(* IEC 61131-3 sources: NachHouse_TST/OSCAT_BasicLib/OscatBasicLib_333a (part 6) *)

(* ---- Device_Driver.ST ---- *)
(* @PATH := '\/Engineering\/automation' *)
FUNCTION_BLOCK DRIVER_1
(*
  driver_1 is a multi purpose driver.
  a rising edge on in sets the output high if toggle is flase. while toggle is true, a rising edge on in toggles the output Q.
  if a timeout is specified the output q will be reset to false automatically after the timeout has elapsed.
  a asynchronous reset and set will force the output high or low respectively.

  version 1.0 2 jan 2008
  programmer  hugo
  tested by   tobias
*)
  VAR_INPUT //???CONSTANT
    Toggle_Mode : BOOL;
    Timeout : TIME;
  END_VAR
  VAR_INPUT
    SET : BOOL;
    IN : BOOL;
    RST : BOOL;
  END_VAR
  VAR_OUTPUT
    Q : BOOL;
  END_VAR
  VAR
    off : TON;
    edge: BOOL;
  END_VAR

  IF off.Q THEN Q := FALSE; END_IF;
  IF rst THEN
    Q := FALSE;
  ELSIF set THEN
    Q := TRUE;
  ELSIF IN AND NOT edge THEN
    IF toggle_mode THEN q := NOT Q; ELSE q := TRUE; END_IF;
  END_IF;
  edge := in;
  IF timeout > t#0s THEN off(in := Q, PT := Timeout); END_IF;

(* revision history
  hm  2. jan 2008   rev 1.0
    original version
*)
END_FUNCTION_BLOCK

(* @PATH := '\/Engineering\/automation' *)
FUNCTION_BLOCK DRIVER_4
(*
  driver_4 is a 4 channel multi purpose driver.
  a rising edge on in? sets the output Q? high if toggle_mode is flase. while toggle_mode is true, a rising edge on in? toggles the output Q?.
  if a timeout is specified the output Q? will be reset to false automatically after the timeout has elapsed.
  a asynchronous reset and set will force the output high or low respectively.
  an asynchronous set will force all outputs high simultaneously

  version 1.0 2 jan 2008
  programmer  hugo
  tested by   tobias
*)
  VAR_INPUT //???CONSTANT
    Toggle_Mode : BOOL;
    Timeout : TIME;
  END_VAR
  VAR_INPUT
    SET : BOOL;
    IN0, IN1, IN2, IN3 : BOOL;
    RST : BOOL;
  END_VAR
  VAR_OUTPUT
    Q0, Q1, Q2, Q3 : BOOL;
  END_VAR
  VAR
    d0, d1, d2, d3 : DRIVER_1;
  END_VAR

  D0(Set:=set, in:=in0, rst:=rst, toggle_mode:=toggle_mode, timeout:=timeout);
  D1(Set:=set, in:=in1, rst:=rst, toggle_mode:=toggle_mode, timeout:=timeout);
  D2(Set:=set, in:=in2, rst:=rst, toggle_mode:=toggle_mode, timeout:=timeout);
  D3(Set:=set, in:=in3, rst:=rst, toggle_mode:=toggle_mode, timeout:=timeout);
  Q0 := D0.Q;
  Q1 := D1.Q;
  Q2 := D2.Q;
  Q3 := D3.Q;

(* revision history
  hm  2. jan 2008   rev 1.0
    original version
*)
END_FUNCTION_BLOCK

(* @PATH := '\/Engineering\/automation' *)
FUNCTION_BLOCK DRIVER_4C
(*
  driver_4C is a multi purpose driver.
  a rising edge on in switches from S0 state S1 and the next edge to state S2 and so on.
  in state S0 all outputs Q are FALSE.
  The stet of the Outputs in any state S? is configurable with setup variables.
  The variables S1..S5 define the states, while the sequence is terminated when a state Variable S? = 0.
  The lower bits 0..3 of the state vars S? are corresponding to the Outputs Q0..Q3

  version 1.0 23. mar. 2009
  programmer  hugo
  tested by tobias
*)
  VAR_INPUT
    IN : BOOL;
    RST : BOOL;
  END_VAR
  VAR_INPUT //??? CONSTANT
    Timeout : TIME;
    SX : ARRAY[1..7] OF BYTE := [1,3,7,15];
  END_VAR
  VAR_OUTPUT
    SN : INT;
    Q0 : BOOL;
    Q1 : BOOL;
    Q2 : BOOL;
    Q3 : BOOL;
  END_VAR
  VAR
    off : TON;
    edge: BOOL;
  END_VAR

  IF RST OR off.Q THEN
    SN := 0;
  ELSIF IN AND NOT edge THEN
    SN := SN + 1;
    IF SN > 7 OR SX[SN] = 0 THEN SN := 0; END_IF;
  END_IF;
  edge := in;
  IF SN > 0 THEN
    Q0 := SX[SN].0;
    Q1 := SX[SN].1;
    Q2 := SX[SN].2;
    Q3 := SX[SN].3;
  ELSE
    Q0 := FALSE;
    Q1 := FALSE;
    Q2 := FALSE;
    Q3 := FALSE;
  END_IF;

  (* maximaum timeout *)
  IF timeout > t#0s THEN off(in := SN > 0, PT := Timeout); END_IF;

(* revision history
  hm  23. mar. 2009 rev 1.0
    original version
*)
END_FUNCTION_BLOCK

(* @PATH := '\/Engineering\/automation' *)
FUNCTION_BLOCK FLOW_CONTROL
(*
  FLOW_CONTROL switches a valves depending on the input in.
  flow control also limits the maximum ontime of the valve and controls pressure on the output side.

  version 1.0 28. jun. 2008
  programmer  hugo
  tested by oscat
*)
  VAR_INPUT
    IN : BOOL;
    REQ : BOOL;
    ENQ : BOOL;
    RST : BOOL;
  END_VAR
  VAR_INPUT //???CONSTANT
    T_AUTO : TIME := T#1h;
    T_DELAY : TIME := T#23h;
  END_VAR
  VAR_OUTPUT
    Q : BOOL;
    STATUS : BYTE;
  END_VAR
  VAR
    timer : TP_1D;
  END_VAR

  STATUS := 100;
  IF RST THEN
    Q := FALSE;
    timer(rst := TRUE);
    timer.RST := FALSE;
    STATUS := 103;
  ELSIF ENQ THEN
    IF IN THEN
      status := 101;
    END_IF;
    IF REQ THEN
      (* timer will generate a timed pulse after TP goes high *)
      timer.PT1 := T_AUTO;
      timer.PTD := T_DELAY;
      timer.IN := TRUE;
      STATUS := 102;
    END_IF;
  END_IF;

  (* set output and run timer *)
  timer();
  timer.IN := FALSE;
  Q := (IN AND ENQ) OR timer.Q;

(* revision history
  hm  28. jun. 2008   rev 1.0
    original version
*)
END_FUNCTION_BLOCK

(* @PATH := '\/Engineering\/automation' *)
FUNCTION_BLOCK FT_Profile
(*
  FT_Profile generates an output signal which is defined by values over a time scale.
  the different values are connected by ramps between the individual values.
  a rising edge on E starts the output signal generation and E = True can delay time_3 / value_3 as long as it stays true.
  an additional multiplier K can be used to multiply the output and an offset O can be added to the output dynamically.

  version 1.1 15 sep 2007
  programmer  tobias
  tested by   hugo
*)
  VAR_INPUT
    K : REAL := 1.0;
    O : REAL;
    M : REAL := 1.0;
    E : BOOL;
  END_VAR
  VAR_INPUT //???CONSTANT
    value_0 : REAL;
    time_1 : TIME;
    value_1 : REAL;
    time_2 : TIME;
    value_2 : REAL;
    time_3 : TIME;
    value_3 : REAL;
    time_10 : TIME;
    value_10 : REAL;
    time_11 : TIME;
    value_11 : REAL;
    time_12 : TIME;
    value_12 : REAL;
    time_13 : TIME;
    value_13 : REAL;
  END_VAR
  VAR_OUTPUT
    Y : REAL;
    RUN : BOOL;
    ET : TIME;
  END_VAR
  VAR
    tx : TIME;
    edge : BOOL;
    state: BYTE;
    ta: TIME;
    tb: TIME;
    t0 : TIME;
    temp: REAL;
    va: REAL;
    vb: REAL;
  END_VAR

  (* read system time *)
  tx := DWORD_TO_TIME(T_PLC_MS());

  (* determine start condition *)
  IF E AND NOT edge THEN
    RUN := TRUE;
    ET := t#0s;
    t0 := tx;
    ta := tx;
    tb := multime(time_1, M);
    va := value_0;
    vb := value_1;
    temp := value_0;
    state := 1;
  END_IF;
  edge := E;

  (* generate startup profile *)
  IF run THEN
    CASE BYTE_TO_USINT(state) OF
      1:  IF tx - ta >= tb THEN
          ta := ta + tb;
          tb := multime(time_2 - time_1, M);
          va := value_1;
          vb := value_2;
          temp := value_1;
          state := 2;
        ELSE
          temp := ((vb - va) * TIME_TO_REAL(tx - ta) / TIME_TO_REAL(tb) + va);
        END_IF;
      2:  IF tx - ta >= tb THEN
          ta := ta + tb;
          tb := multime(time_3 - time_2, M);
          va := value_2;
          vb := value_3;
          temp := value_2;
          state := 3;
        ELSE
          temp := ((vb - va) * TIME_TO_REAL(tx - ta) / TIME_TO_REAL(tb) + va);
        END_IF;
      3:  IF tx - ta >= tb THEN
          ta := ta + tb;
          tb := multime(time_10 - time_3, M);
          va := value_3;
          vb := value_10;
          temp := value_3;
          state := 4;
        ELSE
          temp := ((vb - va) * TIME_TO_REAL(tx - ta) / TIME_TO_REAL(tb) + va);
        END_IF;
      4 : IF tx - ta >= tb THEN
          ta := ta + tb;
          tb := multime(time_11 - time_10, M);
          va := value_10;
          vb := value_11;
          temp := value_10;
          IF E THEN state := 5; ELSE state := 6; END_IF;
        ELSE
          temp := ((vb - va) * TIME_TO_REAL(tx - ta) / TIME_TO_REAL(tb) + va);
        END_IF;
      5:  (* extend the signal while E is true *)
        IF E THEN
          ta := tx;
        ELSE
          state := 6;
        END_IF;
      6:  IF tx - ta >= tb THEN
          ta := ta + tb;
          tb := multime(time_12 - time_11, M);
          va := value_11;
          vb := value_12;
          temp := value_11;
          state := 7;
        ELSE
          temp := ((vb - va) * TIME_TO_REAL(tx - ta) / TIME_TO_REAL(tb) + va);
        END_IF;
      7:  IF tx - ta >= tb THEN
          ta := ta + tb;
          tb := multime(time_13 - time_12, M);
          va := value_12;
          vb := value_13;
          temp := value_12;
          state := 8;
        ELSE
          temp := ((vb - va) * TIME_TO_REAL(tx - ta) / TIME_TO_REAL(tb) + va);
        END_IF;
      8:  IF tx - ta >= tb THEN
          temp := value_13;
          run := FALSE;
        ELSE
          temp := ((vb - va) * TIME_TO_REAL(tx - ta) / TIME_TO_REAL(tb) + va);
        END_IF;
    END_CASE;
    Y := temp * K + O;
    ET := tx - t0;
  END_IF;

(* revision history
  hm  27 feb 2007   rev 1.0
    original version

  hm  15. sep2007   rev 1.1
    replaced Time() with T_PLC_MS for compatibility and performance reasons
*)
END_FUNCTION_BLOCK

(* @PATH := '\/Engineering\/automation' *)
FUNCTION_BLOCK INC_DEC
(*
  incremental decoder with quadruple accuracy.
  2 pulses for each channel are created for each directional pulse.

  version 1.0 4 aug 2006
  programmer  oscat
  tested by   oscat
*)
  VAR_INPUT
    CHa : BOOL;
    CHb : BOOL;
    RST : BOOL;
  END_VAR
  VAR_OUTPUT
    dir : BOOL;
    cnt : INT;
  END_VAR
  VAR
    edgea : BOOL;
    clk: BOOL;
    clka: BOOL;
    clkb: BOOL;
    edgeb: BOOL;
    axb: BOOL;
  END_VAR

  axb := cha XOR chb;

  (* create pulses for channel a *)
  clka := cha XOR edgea;
  edgea := cha;

  clkb := chb XOR edgeb;
  edgeb := chb;

  (* create pulses for both channels *)
  clk := clka OR clkb;

  (* set the direction output *)
  IF axb AND clka THEN dir := TRUE; END_IF;
  IF axb AND clkb THEN dir := FALSE; END_IF;

  (* increment or decrement the counter *)
  IF clk AND dir THEN cnt := cnt + 1; END_IF;
  IF clk AND NOT dir THEN cnt := cnt -1; END_IF;

  (* reset the counter if rst active *)
  IF rst THEN cnt := 0; END_IF;

END_FUNCTION_BLOCK

(* @PATH := '\/Engineering\/automation' *)
FUNCTION_BLOCK INTERLOCK
(*
  INTERLOCK has two inputs I1 and I2 which drive the corresponding outputs Q1 and Q2.
  the inputs signals lock each other out and therfore I1 can only drive Q1 when I2 is Low and vice versa.
  The input TL specifies a dead time between two outputs can become active.
  an output can only become active when the other output was not active for the time TL.

  version 1.0 28 sep 2007
  programmer  hugo
  tested by   tobias
*)
  VAR_INPUT
    I1, I2 : BOOL;
    TL : TIME;
  END_VAR
  VAR_OUTPUT
    Q1, Q2 : BOOL;
  END_VAR
  VAR
    T1, T2 : TOF;
  END_VAR

  (* the input signal have a run delay to lockout the other input *)
  T1(IN := I1, PT := TL);
  T2(IN := I2, PT := TL);

  Q1 := I1 AND NOT t2.Q;
  Q2 := I2 AND NOT t1.Q;

(* revision history
  hm  28 sep 2007   rev 1.0
    original version
*)
END_FUNCTION_BLOCK

(* @PATH := '\/Engineering\/automation' *)
FUNCTION_BLOCK INTERLOCK_4
(*
  INTERLOCK_4 detects one of 4 switches and delivers the number of the switch pressed on the output out
  a output tp is true for one cycle if the output has changed.
  a setup variable MODE selects between 3 different modes:
  MODE = 0, any input active will disable all other inputs
  MODE = 1, the input with the highest number will be acepted
  mode = 2, the input last pressed will disable all others

  version 1.1 14. mar. 2009
  programmer  hugo
  tested by   oscat
*)
  VAR_INPUT
    I0 : BOOL;
    I1 : BOOL;
    I2 : BOOL;
    I3 : BOOL;
    E : BOOL;
    MODE : INT;
  END_VAR
  VAR_OUTPUT
    OUT : BYTE;
    TP : BOOL;
  END_VAR
  VAR
    in: BYTE;
    last: BYTE;
    old: BYTE;
    lmode: INT;
  END_VAR

  (* check if enable is active *)
  IF E THEN
  (* reset all vars when there is a mode change on thy fly *)
    IF mode <> lmode THEN
      out := 0;
      last := 0;
      old := 0;
      lmode := mode;
    END_IF;
    (* load inputs into in *)
    in.0 := I0;
    in.1 := I1;
    in.2 := I2;
    in.3 := I3;
    (* only execute when there is any change *)
    IF in <> last THEN
      (* only execute when inputs have chages state *)
      CASE mode OF
        0:  (* output directly display inputs as bits in byte out *)
          out := in;

        1:  (* the input with the highest number will be acepted *)
          IF in.3 THEN out := 8;
          ELSIF in.2 THEN out := 4;
          ELSIF in.1 THEN out := 2;
          ELSE out := in;
          END_IF;

        2:  (* input last pressed will be displayed only *)
          last := ((in XOR last) AND in);
          IF last.3 THEN out := 8;
          ELSIF last.2 THEN out := 4;
          ELSIF last.1 THEN out := 2;
          ELSE out := last;
          END_IF;

        3:  (* any input active will disable all other inputs *)
          IF (out AND in) = 0 THEN
            IF in.3 THEN out := 8;
            ELSIF in.2 THEN out := 4;
            ELSIF in.1 THEN out := 2;
            ELSE out := in;
            END_IF;
          END_IF;

      END_CASE;
      last := in;
    END_IF;
    tp := out <> old;
    old := out;
  ELSE
    out := 0;
    last := 0;
    old := 0;
    lmode := 0;
    tp := FALSE;
  END_IF;

(* revision history
  hm  24. oct 2008  rev 1.0
    original version

  hm  14. mar. 2009 rev 1.1
    replaced double assignments
*)
END_FUNCTION_BLOCK

(* @PATH := '\/Engineering\/automation' *)
FUNCTION MANUAL : BOOL
(*
  MANUAL is a manual override for digital signals.
  when on and off = FALSE, the output follows IN.
  ON = TRUE forces the output high, and OFF = TRUE forces the output low.

  version 1.0 21. nov. 2008
  programmer  hugo
  tested by oscat
*)
  VAR_INPUT
    IN : BOOL;
    ON : BOOL;
    OFF : BOOL;
  END_VAR

  MANUAL := NOT OFF AND (IN OR ON);

(* revision history
  hm  21. nov 2008  rev 1.0
    original version
*)
END_FUNCTION

(* @PATH := '\/Engineering\/automation' *)
FUNCTION_BLOCK MANUAL_1
(*
  MANUAL_1 is a manual override for digital signals.
  When MAN = FALSE, the output follows IN and when MAN = TRUE the Output follows M_I.

  version 1.2 14. mar. 2009
  programmer  hugo
  tested by   oscat
*)
  VAR_INPUT
    IN : BOOL;
    MAN : BOOL;
    M_I : BOOL;
    SET : BOOL;
    RST : BOOL;
  END_VAR
  VAR_OUTPUT
    Q : BOOL;
    STATUS : BYTE;
  END_VAR
  VAR
    S_edge : BOOL;
    Redge : BOOL;
    edge: BOOL;
  END_VAR

  IF NOT man THEN
    Q := IN;
    STATUS := 100;
    edge := FALSE;
  ELSIF NOT s_edge AND set THEN
    Q := TRUE;
    edge := TRUE;
    status := 101;
  ELSIF NOT Redge AND rst THEN
    Q := FALSE;
    edge := TRUE;
    status := 102;
  ELSIF NOT edge THEN
    Q := M_I;
    status := 103;
  END_IF;

  (* remember levels of manual signals *)
  s_edge := SET;
  Redge := RST;

(* revision history
  hm  17. jun 2008  rev 1.0
    original version

  hm  17. oct 2008  rev 1.1
    deleted unnecessary variable m_edge

  hm  14. mar. 2009 rev 1.2
    replaced double assignments
*)
END_FUNCTION_BLOCK

(* @PATH := '\/Engineering\/automation' *)
FUNCTION_BLOCK MANUAL_2
(*
  MANUAL_2 is a manual override for boolean signals.
  it has static force high and low as well as a manual input.

  version 1.0 22. sep. 2008
  programmer  hugo
  tested by oscat
*)
  VAR_INPUT
    IN : BOOL;
    ENA : BOOL;
    ON : BOOL;
    OFF : BOOL;
    MAN : BOOL;
  END_VAR
  VAR_OUTPUT
    Q : BOOL;
    STATUS : BYTE;
  END_VAR

  IF ena THEN
    IF NOT ON AND NOT OFF THEN
      Q := IN;
      STATUS := 100;
    ELSIF on AND NOT off THEN
      Q := TRUE;
      STATUS := 101;
    ELSIF NOT on AND off THEN
      q := FALSE;
      STATUS := 102;
    ELSE
      Q := MAN;
      STATUS := 103;
    END_IF;
  ELSE
    Q := FALSE;
    STATUS := 104;
  END_IF;

(* revision history
  hm  22. sep. 2008   rev 1.0
    original version
*)
END_FUNCTION_BLOCK

(* @PATH := '\/Engineering\/automation' *)
FUNCTION_BLOCK MANUAL_4
(*
  MANUAL_4 is a manual override for digital signals.
  When MAN = FALSE, the output follows IN and when MAN = TRUE the Output follows M_I.

  version 1.0 17. jun 2008
  programmer  hugo
  tested by oscat
*)
  VAR_INPUT
    I0, I1, I2, I3 : BOOL;
    MAN : BOOL;
    STP : BOOL;
    M0, M1, M2, M3 : BOOL;
  END_VAR
  VAR_OUTPUT
    Q0, Q1, Q2, Q3 : BOOL;
    STATUS : BYTE;
  END_VAR
  VAR
    edge: BOOL;
    pos : INT;
    tog: BOOL;
  END_VAR

  IF man THEN
    IF NOT TOG THEN
      Q0 := M0;
      Q1 := M1;
      Q2 := M2;
      Q3 := M3;
      STATUS := 101;
    END_IF;
    IF STP AND NOT edge THEN
      tog := TRUE;
      CASE pos OF
        0:  Q0 := TRUE;
          Q1 := FALSE;
          Q2 := FALSE;
          Q3 := FALSE;
          STATUS := 110;
        1:  Q0 := FALSE;
          Q1 := TRUE;
          Q2 := FALSE;
          Q3 := FALSE;
          STATUS := 111;
        2:  Q0 := FALSE;
          Q1 := FALSE;
          Q2 := TRUE;
          Q3 := FALSE;
          STATUS := 112;
        3:  Q0 := FALSE;
          Q1 := FALSE;
          Q2 := FALSE;
          Q3 := TRUE;
          STATUS := 113;
      END_CASE;
      pos := INC(pos,1,3);
    END_IF;
  ELSE
    Q0 := I0;
    Q1 := I1;
    Q2 := I2;
    Q3 := I3;
    STATUS := 100;
    tog := FALSE;
    pos := 0;
  END_IF;

  (* remember status of stp *)
  edge := STP;

(* revision history
  hm  17. jun 2008    rev 1.0
    original version
*)
END_FUNCTION_BLOCK

(* @PATH := '\/Engineering\/automation' *)
FUNCTION_BLOCK PARSET
(*
  parset selects on of 4 parameter sets adressed by the inputs A0 and A1. if TC is specified, the change of the outputs
  is ramped by the time tc

  version 1.1 16. mar. 2008
  programmer  hugo
  tested by   tobias
*)
  VAR_INPUT
    A0, A1 : BOOL;
  END_VAR
  VAR_INPUT //???CONSTANT
    X01, X02, X03, X04 : REAL;
    X11, X12, X13, X14 : REAL;
    X21, X22, X23, X24 : REAL;
    X31, X32, X33, X34 : REAL;
    TC : TIME;
  END_VAR
  VAR_OUTPUT
    P1, P2, P3, P4 : REAL;
  END_VAR
  VAR
    X : ARRAY[0..3,1..4] OF REAL;
    S1, S2, S3, S4 : REAL;
    tx, last : UDINT; //DWORD;
    start : BOOL;
    set : USINT; //BYTE;
    init: BOOL;
  END_VAR

  (* read system_time *)
  tx := DWORD_TO_UDINT( T_PLC_MS());

  (* init sequence *)
  IF NOT init THEN
    set.0 := NOT A0;
    init := TRUE;
    X[0,1] := X01;
    X[0,2] := X02;
    X[0,3] := X03;
    X[0,4] := X04;
    X[1,1] := X11;
    X[1,2] := X12;
    X[1,3] := X13;
    X[1,4] := X14;
    X[2,1] := X21;
    X[2,2] := X22;
    X[2,3] := X23;
    X[2,4] := X24;
    X[3,1] := X31;
    X[3,2] := X32;
    X[3,3] := X33;
    X[3,4] := X34;
    P1 := X01;
    P2 := X02;
    P3 := X03;
    P4 := X04;
  END_IF;

  (* check for input change *)
  IF (A0 XOR set.0) OR (A1 XOR set.1) THEN
    (* a new set is selected *)
    set.0 := A0;
    set.1 := A1;
    IF tc > t#0s THEN
      start := TRUE;
      last := tx;
      (* save the step speed for the output changes in S *)
      S1 := (X[set,1] - P1)/DWORD_TO_REAL(TIME_TO_DWORD(tc));
      S2 := (X[set,2] - P2)/DWORD_TO_REAL(TIME_TO_DWORD(tc));
      S3 := (X[set,3] - P3)/DWORD_TO_REAL(TIME_TO_DWORD(tc));
      S4 := (X[set,4] - P4)/DWORD_TO_REAL(TIME_TO_DWORD(tc));
    END_IF;
  ELSIF start AND (tx - last < TIME_TO_UDINT(tc)) THEN
    (* ramp the outputs to the new value *)
    P1 := X[set,1] - S1 * UDINT_TO_REAL(TIME_TO_UDINT(Tc) - tx + last);
    P2 := X[set,2] - S2 * UDINT_TO_REAL(TIME_TO_UDINT(Tc) - tx + last);
    P3 := X[set,3] - S3 * UDINT_TO_REAL(TIME_TO_UDINT(Tc) - tx + last);
    P4 := X[set,4] - S4 * UDINT_TO_REAL(TIME_TO_UDINT(Tc) - tx + last);
  ELSE
    (* make sure outputs match the correct set values *)
    start := FALSE;
    P1 := X[set,1];
    P2 := X[set,2];
    P3 := X[set,3];
    P4 := X[set,4];
  END_IF;

(* revision history
  hm  2.11.2007   rev 1.0
    original version

  hm  16. mar. 2008 rev 1.1
    added type conversions to avoid warnings under codesys 3.0
*)
END_FUNCTION_BLOCK

(* @PATH := '\/Engineering\/automation' *)
FUNCTION_BLOCK PARSET2
(*
  parset2 selects on of 4 parameter sets depending on the value of X. if TC is specified, the change of the outputs
  is ramped by the time TC

  version 1.0 3 nov 2007
  programmer  hugo
  tested by tobias
*)
  VAR_INPUT
    X : REAL;
  END_VAR
  VAR_INPUT //???CONSTANT
    X01, X02, X03, X04 : REAL;
    X11, X12, X13, X14 : REAL;
    X21, X22, X23, X24 : REAL;
    X31, X32, X33, X34 : REAL;
    L1, L2, L3 : REAL;
    TC : TIME;
  END_VAR
  VAR_OUTPUT
    P1,P2,P3,P4 : REAL;
  END_VAR
  VAR
    Pset : parset;
    init: BOOL;
  END_VAR

  (* init sequence *)
  IF NOT init THEN
    init := TRUE;
    pset(TC:=TC, X01:=X01, X02:=X02, X03:=X03, X04:=X04, X11:=X11, X12:=X12, X13:=X13, X14:=X14, X21:=X21, X22:=X22, X23:=X23, X24:=X24, X31:=X31, X32:=X32, X33:=X33, X34:=X34);
  END_IF;
  IF ABS(X) < L1 THEN
    pset(A0 := FALSE, A1 := FALSE);
  ELSIF ABS(X) < L2 THEN
    pset(A0 := TRUE, A1 := FALSE);
  ELSIF ABS(x) < L3 THEN
    pset(A0 := FALSE, A1 := TRUE);
  ELSE
    pset(A0 := TRUE, A1 := TRUE);
  END_IF;
  P1 := pset.P1;
  P2 := pset.P2;
  P3 := pset.P3;
  P4 := pset.P4;

(* revision history
  hm    3.11.2007   rev 1.0
    original version
*)
END_FUNCTION_BLOCK

(* @PATH := '\/Engineering\/automation' *)
FUNCTION_BLOCK SIGNAL
(*
  this function generates an output signal according to a bit pattern SIG.
  the patter is shifted to the output in time steps of TS.
  ts defaults to 128 ms if not specified.

  version 1.0 13 dec 2007
  programmer  hugo
  tested by   tobias
*)
  VAR_INPUT
    IN : BOOL;
    SIG : BYTE;
    TS : TIME;
  END_VAR
  VAR_OUTPUT
    Q : BOOL;
  END_VAR
  VAR
    tx: UDINT; //DWORD;
    step: BYTE;
  END_VAR
  VAR CONSTANT
    one : BYTE := 1;
  END_VAR

  IF in THEN
    (* an alarm is present read system time first *)
    tx := DWORD_TO_UDINT( T_PLC_MS());
    (* calculate the step counter which is the lowest 3 bits of (time / ts) *)
    IF ts > t#0s THEN
      step := DWORD_TO_BYTE( UDINT_TO_DWORD(tx / TIME_TO_UDINT(ts)) AND 16#0000_0007);
    ELSE
      step := DWORD_TO_BYTE(SHR( UDINT_TO_DWORD(tx),7) AND 16#0000_0007);
    END_IF;
    (* convert the value 0-7 in step into one bit only (bit 0-7) *)
    step := SHL(one,BYTE_TO_UINT(step));
    (* generate the output signal *)
    Q := (step AND sig) > 0;
  ELSE
    Q := FALSE;
  END_IF;

(* revision history
  hm  13.12.2007    rev 1.0
    original version
*)
END_FUNCTION_BLOCK

(* @PATH := '\/Engineering\/automation' *)
FUNCTION_BLOCK SIGNAL_4
(*
  this function generates one out of 4 signals specified by bit patterns S1 .. S4.
  the selected pattern will be shifted with the step time TS.
  In1 has higher priority then In2 which has higher priority then IN3 and in4 has the lowest priority.
  ts defaults to 128 ms if not specified.

  version 1.0 13 dec 2007
  programmer  hugo
  tested by   tobias
*)
  VAR_INPUT
    IN1 : BOOL;
    IN2 : BOOL;
    IN3 : BOOL;
    IN4 : BOOL;
    TS : TIME;
  END_VAR
  VAR_INPUT //???CONSTANT
    S1 : BYTE := 2#1111_1111;
    S2 : BYTE := 2#1111_0000;
    S3 : BYTE := 2#1010_1010;
    S4 : BYTE := 2#1010_0000;
  END_VAR
  VAR_OUTPUT
    Q : BOOL;
  END_VAR
  VAR
    sig : SIGNAL;
  END_VAR

  (* an alarm is present read system time first *)
  (* check if an alarm is present if yes set sig to the alarm pattern otherwise exit the routine *)
  IF in1 THEN
    sig(in := TRUE, sig := s1, TS := TS);
  ELSIF in2 THEN
    sig(in := TRUE, sig := s2, TS := TS);
  ELSIF in3 THEN
    sig(in := TRUE, sig := s3, TS := TS);
  ELSIF in4 THEN
    sig(in := TRUE, sig := s4, TS := TS);
  ELSE
    sig(in := FALSE);
  END_IF;

  (* set the output *)
  Q := sig.Q;

(* revision history
  hm  13.12.2007    rev 1.0
    original version
*)
END_FUNCTION_BLOCK

(* @PATH := '\/Engineering\/automation' *)
FUNCTION_BLOCK SRAMP
(*
  RAMPS generates output signal which are slew rate and acceleration controlled.

  version 1.1 11. mar. 2009
  programmer  hugo
  tested by   tobias
*)
  VAR_INPUT
    X : REAL;
    A_UP : REAL;
    A_DN :REAL;
    VU_MAX : REAL;
    VD_MAX : REAL;
    LIMIT_HIGH : REAL;
    LIMIT_LOW : REAL;
    RST : BOOL;
  END_VAR
  VAR_OUTPUT
    Y : REAL;
    V : REAL;
  END_VAR
  VAR
    cycle_time : TC_S;
    init: BOOL;
  END_VAR

  (* read the system_time in microseconds *)
  cycle_time();

  (* assure range of inputs *)
  A_up := MAX(0.0, A_UP);
  A_dn := MIN(0.0, A_dn);
  VU_max := MAX(0.0, VU_max);
  VD_max := MIN(0.0, VD_MAX);

  (* calculate the output offset *)
  IF rst OR NOT init THEN
    init := TRUE;
    Y := 0.0;
    V := 0.0;
  ELSIF X = Y THEN
    v := 0.0;
  ELSIF X > Y THEN
    (* output is too low >> ramp up and brake at the end *)
    (* accelerate the speed and limit to vu_max *)
    v := MIN(v + A_UP * cycle_time.TC, vu_max);
    (* calculate the max speed to be able to brake and select the lowest *)
    v := MIN(SQRT((Y-X) * 2.0 * A_DN), v);
    (* calculate the output and obey limits *)
    y := LIMIT(limit_low, y + MIN(v * cycle_time.TC, X-Y), limit_high);
  ELSIF X < Y THEN
    (* output is too high >> ramp dn and brake at the end *)
    (* accelerate the speed and limit to vd_max *)
    v := MAX(v + A_DN * cycle_time.TC, vd_max);
    (* calculate the max speed to be able to brake and select the lowest *)
    v := MAX(-SQRT((Y-X) * 2.0 * A_UP), v);
    (* calculate the output and obey limits *)
    y := LIMIT(limit_low, y + MAX(v * cycle_time.TC, X-Y), limit_high);
  END_IF;

(* revision history
  hm  13. mar. 2008 rev 1.0
    original version

  hm  11. mar. 2009 rev 1.1
  	real constants updated to new systax using dot
*)
END_FUNCTION_BLOCK

(* @PATH := '\/Engineering\/automation' *)
FUNCTION_BLOCK TUNE
(*
  tune generates an output signal which is set by input switches.
  up to 4 switsches can be used to tune the signal up or down.

  version 1.2 11. mar. 2009
  programmer  hugo
  tested by   tobias
*)
  VAR_INPUT
    SET : BOOL;
    SU, SD : BOOL;
    RST : BOOL;
  END_VAR
  VAR_INPUT //???CONSTANT
    SS : REAL := 0.1;
    Limit_L : REAL;
    LIMIT_H : REAL := 100.0;
    RST_val : REAL;
    SET_val : REAL := 100.0;
    T1 : TIME := T#500ms;
    T2 : TIME := T#2s;
    S1 : REAL := 2.0;
    S2 : REAL := 10.0;
  END_VAR
  VAR_OUTPUT
    Y : REAL;
  END_VAR
  VAR
    tx : UDINT; //DWORD;
    start, start2 : UDINT; //DWORD;
    state : INT;
    in : BOOL;
    step : REAL;
    SPEED : REAL;
    Y_start : REAL;
    Y_start2: REAL;
  END_VAR

  (* read system time *)
  tx := DWORD_TO_UDINT( T_PLC_MS());

  IF rst THEN
    Y := RST_val;
    state := 0;
  ELSIF set THEN
    Y := SET_val;
    state := 0;
  ELSIF state > 0 THEN
    (* key has been pushed state machine operating *)
    (* first read the correct input *)
    IF state = 1 THEN
      (* step up *)
      in := su;
    ELSE
      (* step down *)
      in := sd;
    END_IF;
    (* check for single step operation *)
    IF NOT in AND (tx - start <= TIME_TO_UDINT(T1)) THEN
      Y := Y_start + step;
      state := 0;
    (* check if fast ramp needs to be generated *)
    ELSIF in AND (tx - start >= TIME_TO_UDINT(T2)) THEN
      Y := Y_start2 + UDINT_TO_REAL(tx - start2) * s2 / speed;
    (* check if slow ramp needs to be generated *)
    ELSIF in AND (tx - start >= TIME_TO_UDINT(T1)) THEN
      Y := Y_start + UDINT_TO_REAL(tx - start - TIME_TO_UDINT(T1)) * S1 / speed;
      start2 := tx;
      Y_start2 := Y;
    ELSIF NOT in THEN
      state := 0;
    END_IF;
  ELSIF su THEN
    (* slow step up *)
    state := 1;
    start := tx;
    step := ss;
    speed := 1000.0;
    Y_start := Y;
  ELSIF sd THEN
    (* slow step down *)
    state := 2;
    start := tx;
    step := -ss;
    speed := -1000.0;
    Y_start := Y;
  END_IF;

  (* make sure output does not exceed limits *)
  Y := LIMIT(LIMIT_L, Y, LIMIT_H);

(* revision history
  hm  3.11.2007   rev 1.0
    original version

  hm  16. mar. 2008 rev 1.1
    added type conversions to avoid warnings under codesys 3.0

  hm  11. mar. 2009 rev 1.2
  	real constants updated to new systax using dot
*)
END_FUNCTION_BLOCK

(* @PATH := '\/Engineering\/automation' *)
FUNCTION_BLOCK TUNE2
(*
  tune2 generates an output signal which is set by input switches.
  up to 4 switsches can be used to tune the signal up or down.

  version 1.2 11. mar. 2009
  programmer  hugo
  tested by   tobias
*)
  VAR_INPUT
    SET : BOOL;
    SU, SD : BOOL;
    FU, FD : BOOL;
    RST : BOOL;
  END_VAR
  VAR_INPUT //???CONSTANT
    SS : REAL := 0.1;
    FS : REAL := 5.0;
    Limit_L : REAL;
    LIMIT_H : REAL := 100.0;
    RST_val : REAL;
    SET_val : REAL := 100.0;
    TR : TIME := T#500ms;
    S1 : REAL := 2.0;
    S2 : REAL := 10.0;
  END_VAR
  VAR_OUTPUT
    Y : REAL;
  END_VAR
  VAR
    tx : UDINT; //DWORD;
    start : UDINT; //DWORD;
    state : INT;
    in : BOOL;
    step : REAL;
    SPEED : REAL;
    Y_start : REAL;
  END_VAR

  (* read system time *)
  tx := DWORD_TO_UDINT( T_PLC_MS());

  IF rst THEN
    Y := RST_val;
    state := 0;
  ELSIF set THEN
    Y := SET_val;
    state := 0;
  ELSIF state > 0 THEN
    (* key has been pushed state machine operating *)
    (* first read the correct input *)
    CASE state OF
      1 : (* slow up *)
        in := su;
      2 : (* slow down *)
        in := sd;
      3 : (* fast up *)
        in := fu;
      4 : (* fast down *)
        in := fd;
    END_CASE;
    (* check for single step operation *)
    IF NOT in AND (tx - start <= TIME_TO_UDINT(TR)) THEN
      Y := Y_start + step;
      state := 0;
    (* check if ramp needs to be generated *)
    ELSIF in AND (tx - start >= TIME_TO_UDINT(TR)) THEN
      Y := Y_start + UDINT_TO_REAL(tx - start - TIME_TO_UDINT(TR)) * speed;
    ELSIF NOT in THEN
      state := 0;
    END_IF;
  ELSIF su THEN
    (* slow step up *)
    state := 1;
    start := tx;
    step := ss;
    speed := s1 * 1.0E-3;
    Y_start := Y;
  ELSIF sd THEN
    (* slow step down *)
    state := 2;
    start := tx;
    step := -ss;
    speed := -s1 * 1.0E-3;
    Y_start := Y;
  ELSIF fu THEN
    (* fast step up *)
    state := 3;
    start := tx;
    step := fs;
    speed := s2 * 1.0E-3;
    y_start := Y;
  ELSIF fd THEN
    (* fast step down *)
    state := 4;
    start := tx;
    step := -fs;
    speed := -s2 * 1.0E-3;
    y_start := Y;
  END_IF;

  (* make sure output does not exceed limits *)
  Y := LIMIT(LIMIT_L, Y, LIMIT_H);

(* revision history
  hm  3.11.2007   rev 1.0
    original version

  hm  16. 3. 2008 rev 1.1
    added type conversions to avoid warnings in codesys 3.0
    improved performance

  hm  11. mar. 2009 rev 1.2
  	real constants updated to new systax using dot
*)
END_FUNCTION_BLOCK

(* ---- Latches_FlipFlop_ShiftRegister.ST ---- *)
(* @PATH := '\/Logic\/FF edge triggered' *)
FUNCTION_BLOCK COUNT_BR
(*
  Count_BR is a byte counter with independen up and dn inputs. the counter counts from 0 to mx and continues at 0 after is has reached mx
  a step input sets the counters stepping width.

  version 1.0 16 jan 2008
  programmer  hugo
  tested BY tobias
*)
  VAR_INPUT
    SET : BOOL;
    IN : BYTE;
    UP : BOOL;
    DN : BOOL;
    STEP : BYTE := 1;
    MX : BYTE := 255;
    RST : BOOL;
  END_VAR
  VAR_OUTPUT
    CNT : BYTE;
  END_VAR
  VAR
    last_up: BOOL;
    last_dn: BOOL;
  END_VAR

  IF rst THEN
    cnt := 0;
  ELSIF set THEN
    cnt := LIMIT(0,in,mx);
  ELSIF up AND NOT last_up THEN
    cnt := INT_TO_BYTE(INC( BYTE_TO_INT(cnt),BYTE_TO_INT(step),BYTE_TO_INT(mx)));
  ELSIF dn AND NOT last_dn THEN
    cnt := INT_TO_BYTE(INC( BYTE_TO_INT(cnt),-BYTE_TO_INT(step),BYTE_TO_INT(mx)));
  END_IF;
  last_up := up;
  last_dn := dn;

(* revision history
  hm  16. jan 2008  rev 1.0
    original version
*)
END_FUNCTION_BLOCK

(* @PATH := '\/Logic\/FF edge triggered' *)
FUNCTION_BLOCK COUNT_DR
(*
  Count_DR is a DWORD counter with independen up and dn inputs. the counter counts from 0 to mx and continues at 0 after is has reached mx
  a step input sets the counters stepping width.

  version 1.1 20. jan. 2011
  programmer  hugo
  tested BY   tobias
*)
  VAR_INPUT
    SET : BOOL;
    IN : DWORD;
    UP : BOOL;
    DN : BOOL;
    STEP : DWORD := 1;
    MX : DWORD := 16#FFFFFFFF;
    RST : BOOL;
  END_VAR
  VAR_OUTPUT
    CNT : DWORD;
  END_VAR
  VAR
    last_up: BOOL;
    last_dn: BOOL;
  END_VAR

  IF rst THEN
    cnt := 0;
  ELSIF set THEN
    cnt := LIMIT(0,in,mx);
  ELSIF up AND NOT last_up THEN
    IF STEP > UDINT_TO_DWORD( DWORD_TO_UDINT(MX) - DWORD_TO_UDINT(CNT)) THEN
      CNT := UDINT_TO_DWORD( DWORD_TO_UDINT(CNT) - DWORD_TO_UDINT(MX) + DWORD_TO_UDINT(STEP) - 1);
    ELSE
      CNT := UDINT_TO_DWORD( DWORD_TO_UDINT(CNT) + DWORD_TO_UDINT(STEP));
    END_IF;
  ELSIF dn AND NOT last_dn THEN
    IF STEP > CNT THEN
      CNT := UDINT_TO_DWORD( DWORD_TO_UDINT(CNT) - DWORD_TO_UDINT(STEP) + DWORD_TO_UDINT(MX) + 1);
    ELSE
      CNT := UDINT_TO_DWORD( DWORD_TO_UDINT(CNT) - DWORD_TO_UDINT(STEP));
    END_IF;
  END_IF;
  last_up := up;
  last_dn := dn;

(* revision history
  hm  12. jun 2008  rev 1.0
    original version

  hm  20. jan. 2011 rev 1.1
    corrected init value of MX to 16#FFFFFFFF
*)
END_FUNCTION_BLOCK

(* @PATH := '\/Logic\/FF edge triggered' *)
FUNCTION_BLOCK FF_D2E
(*
  dual D-type flip flop with reset and rising clock trigger

  version 1.3 14. mar. 2009
  programmer  hugo
  tested by   oscat
*)
  VAR_INPUT
    D0 : BOOL;
    D1 : BOOL;
    CLK : BOOL;
    RST : BOOL;
  END_VAR
  VAR_OUTPUT
    Q0 : BOOL;
    Q1 : BOOL;
  END_VAR
  VAR
    edge : BOOL;
  END_VAR

  IF rst THEN
    Q0 := FALSE;
    Q1 := FALSE;
  ELSIF clk AND NOT edge THEN
    Q0 := D0;
    Q1 := D1;
  END_IF;
  edge := CLK;

(* revision history
  hm  25. dec 2007  rev 1.0
    original version

  hm  27. dec 2007  rev 1.1
    changed code for better performance

  hm  30. oct. 200  rev 1.2
    deleted unnecessary init with 0

  hm  14. mar. 2009 rev 1.3
    removed double assignments
*)
END_FUNCTION_BLOCK

(* @PATH := '\/Logic\/FF edge triggered' *)
FUNCTION_BLOCK FF_D4E
(*
  quad D-type flip flop with reset and rising clock trigger

  version 1.3 14. mar. 2009
  programmer  hugo
  tested by   oscat
*)
  VAR_INPUT
    D0 : BOOL;
    D1 : BOOL;
    D2 : BOOL;
    D3 : BOOL;
    CLK : BOOL;
    RST : BOOL;
  END_VAR
  VAR_OUTPUT
    Q0 : BOOL;
    Q1 : BOOL;
    Q2 : BOOL;
    Q3 : BOOL;
  END_VAR
  VAR
    edge : BOOL;
  END_VAR

  IF rst THEN
    Q0 := FALSE;
    Q1 := FALSE;
    Q2 := FALSE;
    Q3 := FALSE;
  ELSIF clk AND NOT edge THEN
    Q0 := D0;
    Q1 := D1;
    Q2 := D2;
    Q3 := D3;
  END_IF;
  edge := CLK;

(* revision history
  hm  4. aug 2006 rev 1.0
    original version

  hm  27. dec 2007  rev 1.1
    changed code for better performance

  hm  30. oct. 200  rev 1.2
    deleted unnecessary init with 0

  hm  14. mar. 2009 rev 1.3
    removed double assignments
*)
END_FUNCTION_BLOCK

(* @PATH := '\/Logic\/FF edge triggered' *)
FUNCTION_BLOCK FF_DRE
(*
  D-type flip flop with set, reset and rising clock trigger

  version 1.2 30. oct. 2008
  programmer  hugo
  tested by oscat
*)
  VAR_INPUT
    SET : BOOL;
    D : BOOL;
    CLK : BOOL;
    RST : BOOL;
  END_VAR
  VAR_OUTPUT
    Q : BOOL;
  END_VAR
  VAR
    edge : BOOL;
  END_VAR

  IF rst OR set THEN
    Q := NOT rst;
  ELSIF clk AND NOT edge THEN
    Q := D;
  END_IF;
  edge := CLK;

(* revision history
  hm  4. aug 2006   rev 1.0
    original version

  hm  27. dec 2007  rev 1.1
    changed code for better performance

  hm  30. oct. 2008 rev 1.2
    optimized performance
*)
END_FUNCTION_BLOCK

(* @PATH := '\/Logic\/FF edge triggered' *)
FUNCTION_BLOCK FF_JKE
(*
  JK-type flip flop with set, reset and rising clock trigger
  set and reset are asynchron while the FF is rising edge triggered
  J=0 and K=0 and CLK >>> no action
  J=1 and K=0 and CLK >>> output = 1
  J=0 and K=1 and CLK >>> output = 0
  J=1 and K=1 and CLK >>> toggle output

  version 1.2 30. oct. 2008
  programmer  hugo
  tested by oscat
*)
  VAR_INPUT
    SET : BOOL;
    J : BOOL;
    CLK : BOOL;
    K : BOOL;
    RST : BOOL;
  END_VAR
  VAR_OUTPUT
    Q : BOOL;
  END_VAR
  VAR
    edge : BOOL;
  END_VAR

  IF rst OR set THEN
    Q := NOT rst;
  ELSIF clk AND NOT edge THEN
    IF J XOR K THEN Q := J;
    ELSE Q := K XOR Q;
    END_IF;
  END_IF;
  edge := CLK;

(* revision history
  hm  4. aug 2006   rev 1.0
    original version

  hm  27. dec 2007  rev 1.1
    changed code for better performance

  hm  30. oct. 2008 rev 1.2
    optimized performance
*)
END_FUNCTION_BLOCK

(* @PATH := '\/Logic\/FF edge triggered' *)
FUNCTION_BLOCK FF_RSE
(*
  this is a rising edge triggered rs flip flop
  a rising edge on CS sets Q = TRUE and a rising edge on CR sets Q = FALSE.
  CR has priority over CS.

  version 1.0 16. jul. 2008
  programmer  hugo
  tested by oscat
*)
  VAR_INPUT
    CS : BOOL;
    CR : BOOL;
    RST : BOOL;
  END_VAR
  VAR_OUTPUT
    Q : BOOL;
  END_VAR
  VAR
    es, er : BOOL;
  END_VAR

  IF rst THEN
    (* asynchronous reset *)
    Q := FALSE;
  ELSIF CR AND NOT er THEN
    (* rising edge on CR *)
    Q := FALSE;
  ELSIF CS AND NOT es THEN
    (* rising edge on CS *)
    Q := TRUE;
  END_IF;
  es := CS;
  er := CR;

(* revision history
  hm  16. jul. 2008 rev 1.0
    original version
*)
END_FUNCTION_BLOCK

(* @PATH := '\/Logic\/FF edge triggered' *)
FUNCTION_BLOCK SELECT_8
(*
  select_8 selects one of 8 outputs at any time. the outputscan be selected by up or down keys and an independent anable switches all outouts off if set false

  version 1.1 27. feb. 2009
  programmer  hugo
  tested BY   oscat
*)
  VAR_INPUT
    E : BOOL;
    SET : BOOL;
    IN : BYTE;
    UP : BOOL;
    DN : BOOL;
    RST : BOOL;
  END_VAR
  VAR_OUTPUT
    Q0, Q1, Q2, Q3, Q4, Q5, Q6, Q7 : BOOL;
    STATE : INT;
  END_VAR
  VAR
    last_up: BOOL;
    last_dn : BOOL;
  END_VAR

  IF rst THEN
    state := 0;
  ELSIF set THEN
    state := BYTE_TO_INT(IN);
  ELSIF up AND NOT last_up THEN
    state := inc(state,1,7);
  ELSIF dn AND NOT last_dn THEN
    state := inc(state,-1,7);
  END_IF;
  last_UP := UP;
  last_DN := DN;

  Q0 := FALSE;
  Q1 := FALSE;
  Q2 := FALSE;
  Q3 := FALSE;
  Q4 := FALSE;
  Q5 := FALSE;
  Q6 := FALSE;
  Q7 := FALSE;

  IF E THEN
    CASE state OF
      0: Q0 := TRUE;
      1: Q1 := TRUE;
      2: Q2 := TRUE;
      3: Q3 := TRUE;
      4: Q4 := TRUE;
      5: Q5 := TRUE;
      6: Q6 := TRUE;
      7: Q7 := TRUE;
    END_CASE;
  END_IF;

(* revision history
  hm  16. jan 2008  rev 1.0
    original version

  hm  27. feb. 2009 rev 1.1
    renamed input en to e
*)
END_FUNCTION_BLOCK

(* @PATH := '\/Logic\/FF edge triggered' *)
FUNCTION_BLOCK SHR_4E
(*
  4 bit shift register with reset

  version 1.1 25. oct. 2008
  programmer  hugo
  tested by   tobias
*)
  VAR_INPUT
    SET : BOOL;
    D0: BOOL;
    CLK: BOOL;
    RST: BOOL;
  END_VAR
  VAR_OUTPUT
    Q0: BOOL;
    Q1: BOOL;
    Q2: BOOL;
    Q3: BOOL;
  END_VAR
  VAR
    trig : R_TRIG;
  END_VAR

  (* trig.Q signals a rising edge on clk *)
  trig(clk := clk);

  IF set OR rst THEN
    Q0 := NOT rst;
    Q1 := Q0;
    Q2 := Q0;
    Q3 := Q0;
  ELSIF trig.Q THEN
    Q3 := Q2;
    Q2 := Q1;
    Q1 := Q0;
    Q0 := D0;
  END_IF;

(* revision history
  hm  4. aug. 2006  rev 1.0
    original version

  hm  25. oct. 2008 rev 1.1
    optimized code
*)
END_FUNCTION_BLOCK

(* @PATH := '\/Logic\/FF edge triggered' *)
FUNCTION_BLOCK SHR_4UDE
(*
  4 bit shift register with reset up / down direction input

  version 1.2 14. mar. 2009
  programmer  hugo
  tested by   tobias
*)
  VAR_INPUT
    SET : BOOL;
    D0: BOOL;
    D3: BOOL;
    CLK: BOOL;
    DN : BOOL;
    RST: BOOL;

  END_VAR
  VAR_OUTPUT
    Q0: BOOL;
    Q1: BOOL;
    Q2: BOOL;
    Q3: BOOL;
  END_VAR
  VAR
    trig : R_TRIG;
  END_VAR

  (* trig.Q signals a rising edge on clk *)
  trig(clk := clk);

  IF set OR rst THEN
    Q0 := NOT RST;
    Q1 := Q0;
    Q2 := Q0;
    Q3 := Q0;
  ELSIF trig.Q THEN
    IF dn THEN
      Q0 := Q1;
      Q1 := Q2;
      Q2 := Q3;
      Q3 := D3;
    ELSE
      Q3 := Q2;
      Q2 := Q1;
      Q1 := Q0;
      Q0 := D0;
    END_IF;
  END_IF;

(* revision history
  hm  4. aug. 2006  rev 1.0
    original version

  hm  25. oct. 2008 rev 1.1
    optimized code

  hm  14. mar. 2009 rev 1.2
    removed double assignments
*)
END_FUNCTION_BLOCK

(* @PATH := '\/Logic\/FF edge triggered' *)
FUNCTION_BLOCK SHR_8PLE
(*
  8 bit shift register with reset and parallel load
  the register can shift up or down
  it also has a serial input.
  the Din input is on Bit0 for up shift and on bit 7 for down shift
  the Dout output is on Bit7 for up shift and on bit 0 for down shift
  paralle clock is performed clock synchron while a shift is performed first and then the register is reloaded

  version 1.0 4 aug 2006
  programmer  hugo
  tested by oscat
*)
  VAR_INPUT
    Din : BOOL;
    Dload : BYTE;
    CLK: BOOL;
    UP: BOOL :=1;
    load : BOOL;
    RST: BOOL;
  END_VAR
  VAR_OUTPUT
    DOut: BOOL;
  END_VAR
  VAR
    edge : BOOL :=1;
    register : BYTE;
  END_VAR

  (* flankenerkennung clk wird high und edge war high reset ist nicht aktiv und set ist nicht aktiv *)
  IF CLK AND edge AND NOT rst THEN
    edge := FALSE;  (* flanke wurde erkannt und weitere flankenerkennung wird verhindert bis edge wieder true ist *)
    (* hier ist der code für das flankenevent *)
    IF UP THEN            (*shift up *)
      register := SHL(register,1);
      register.0 := Din;
      Dout := register.7;
    ELSE                (* shift down *);
      register := SHR(register,1);
      register.7 := Din;
      Dout := register.0;
    END_IF;
    IF load THEN              (* the byte on Din will be loaded if load = true *)
      register := Dload;
      IF up THEN Dout := register.7; ELSE Dout := register.0; END_IF;
    END_IF;
  END_IF;
  IF NOT clk THEN edge := TRUE; END_IF; (* sobald clk wieder low wird warten auf nächste flanke *)
  IF rst THEN                 (* wenn reset aktiv dann ausgang rücksetzen *)
    register := 0;
    Dout := FALSE;
  END_IF;
END_FUNCTION_BLOCK

(* @PATH := '\/Logic\/FF edge triggered' *)
FUNCTION_BLOCK SHR_8UDE
(*
  8 bit shift register with reset

  version 1.2 14. mar. 2009
  programmer  hugo
  tested by   tobias
*)
  VAR_INPUT
    SET : BOOL;
    D0: BOOL;
    D7: BOOL;
    CLK: BOOL;
    DN : BOOL;
    RST: BOOL;
  END_VAR
  VAR_OUTPUT
    Q0: BOOL;
    Q1: BOOL;
    Q2: BOOL;
    Q3: BOOL;
    Q4: BOOL;
    Q5: BOOL;
    Q6: BOOL;
    Q7: BOOL;
  END_VAR
  VAR
    trig : R_TRIG;
  END_VAR

  (* trig.Q signals a rising edge on clk *)
  trig(clk := clk);

  IF set OR rst THEN
    Q0 := NOT RST;
    Q1 := Q0;
    Q2 := Q0;
    Q3 := Q0;
    Q4 := Q0;
    Q5 := Q0;
    Q6 := Q0;
    Q7 := Q0;
  ELSIF trig.Q THEN
    IF dn THEN
      Q0 := Q1;
      Q1 := Q2;
      Q2 := Q3;
      Q3 := Q4;
      Q4 := Q5;
      Q5 := Q6;
      Q6 := Q7;
      Q7 := D7;
    ELSE
      Q7 := Q6;
      Q6 := Q5;
      Q5 := Q4;
      Q4 := Q3;
      Q3 := Q2;
      Q2 := Q1;
      Q1 := Q0;
      Q0 := D0;
    END_IF;
  END_IF;

(* revision history
  hm  4. aug. 2006  rev 1.0
    original version

  hm  25. oct. 2008 rev 1.1
    optimized code

  hm  14. mar. 2009 rev 1.2
    removed double assignments
*)
END_FUNCTION_BLOCK

(* @PATH := '\/Logic\/FF edge triggered' *)
FUNCTION_BLOCK TOGGLE
(*
  toggle flip flop the output changes state with every rising edge of clk.

  version 1.1 30. oct. 2008
  programmer  hugo
  tested by oscat
*)
  VAR_INPUT
    CLK : BOOL;
    rst : BOOL;
  END_VAR
  VAR_OUTPUT
    Q : BOOL;
  END_VAR
  VAR
    edge : BOOL;
  END_VAR

  IF rst THEN
    q := 0;
  ELSIF clk AND NOT edge THEN
    Q := NOT Q;
  END_IF;
  edge := clk;

(* revision history
  hm  13.9.2007   rev 1.0
    original version

  hm  30. oct. 2008 rev 1.1
    deleted unnecessary init
*)
END_FUNCTION_BLOCK

(* @PATH := '\/Logic\/FF pulse triggered' *)
FUNCTION_BLOCK LTCH
(*
  Transparent Latch with asynchronous reset

  version 1.2 30. oct. 2008
  programmer  hugo
  tested by oscat
*)
  VAR_INPUT
    D : BOOL;
    L : BOOL;
    RST : BOOL;
  END_VAR
  VAR_OUTPUT
    Q : BOOL;
  END_VAR

  (* as long as L is true, the latch is transparent and and change of D is transferred to Q *)
  (* of course only when there is no asynchronous reset *)
  IF rst THEN       (* if asynchronous reset then Q=0 *)
    Q := FALSE;
  ELSIF L THEN      (* latch is transparent *)
    Q := D;
  END_IF;

(* revision history
  hm  4. aug 2006   rev 1.0
    original version

  hm  27. dec 2007  rev 1.1
    changed code for better performance

  hm  30. oct. 2008 rev 1.2
    deleted unnecessary init with 0
*)
END_FUNCTION_BLOCK

(* @PATH := '\/Logic\/FF pulse triggered' *)
FUNCTION_BLOCK LTCH_4
(*
  Quad Transparent Latch with asynchronous reset

  version 1.3 14. mar. 2009
  programmer  hugo
  tested by   oscat
*)
  VAR_INPUT
    D0 : BOOL;
    D1 : BOOL;
    D2 : BOOL;
    D3 : BOOL;
    L : BOOL;
    RST : BOOL;
  END_VAR
  VAR_OUTPUT
    Q0 : BOOL;
    Q1 : BOOL;
    Q2 : BOOL;
    Q3 : BOOL;
  END_VAR

  (* as long as L is true, the latch is transparent and and change of D is transferred to Q *)
  (* of course only when there is no asynchronous reset *)
  IF rst THEN     (* if asynchronous reset then Q=0 *)
    Q0 := FALSE;
    Q1 := FALSE;
    Q2 := FALSE;
    Q3 := FALSE;
  ELSIF L THEN      (* latch is transparent *)
    Q0 := D0;
    Q1 := D1;
    Q2 := D2;
    Q3 := D3;
  END_IF;

(* revision history
  hm  4. aug 2006 rev 1.0
    original version

  hm  27. dec 2007  rev 1.1
    changed code for better performance

  hm  30. oct. 2008 rev 1.2
    deleted unnecessary init with 0

  hm  14. mar. 2009 rev 1.3
    removed double assignments
*)
END_FUNCTION_BLOCK

(* @PATH := '\/Logic\/FF pulse triggered' *)
FUNCTION_BLOCK STORE_8
(*
  Store_4 stores up to 4 boolean inputs until a reset is clearing the outputs.
  the respective output is set with a true at the respective input and stays true until a reset is generated.
  a set input is used to set all outputs true at the same time, independent of their inputs.
  a clear input is used to reset only the lowest priority of the outputs one at a time.
  the lowest priority is q3.

  version 1.2 14. mar. 2009
  programmer  hugo
  tested by   oscat
*)
  VAR_INPUT
    Set : BOOL;
    D0,D1, D2, D3, D4, D5, D6, D7 : BOOL;
    Clr : BOOL;
    Rst : BOOL;
  END_VAR
  VAR_OUTPUT
    Q0, Q1, Q2, Q3, Q4, Q5, Q6, Q7 : BOOL;
  END_VAR
  VAR
    edge: BOOL;
  END_VAR

  IF rst OR set THEN
    q0 := NOT rst;
    q1 := q0;
    q2 := q0;
    q3 := q0;
    q4 := q0;
    q5 := q0;
    q6 := q0;
    q7 := q0;
  ELSE
    IF D0 THEN Q0 := TRUE; END_IF;
    IF D1 THEN Q1 := TRUE; END_IF;
    IF D2 THEN Q2 := TRUE; END_IF;
    IF D3 THEN Q3 := TRUE; END_IF;
    IF D4 THEN Q4 := TRUE; END_IF;
    IF D5 THEN Q5 := TRUE; END_IF;
    IF D6 THEN Q6 := TRUE; END_IF;
    IF D7 THEN Q7 := TRUE; END_IF;

    IF clr AND NOT edge THEN
      IF q0 THEN q0 := FALSE;
      ELSIF q1 THEN q1 := FALSE;
      ELSIF q2 THEN q2 := FALSE;
      ELSIF q3 THEN q3 := FALSE;
      ELSIF q4 THEN q4 := FALSE;
      ELSIF q5 THEN q5 := FALSE;
      ELSIF q6 THEN q6 := FALSE;
      ELSE q7 := FALSE;
      END_IF;
    END_IF;
    edge := clr;
  END_IF;

(* revision history
  hm  25.12.2007  rev 1.0
    original version

  hm  30. oct. 2008 rev 1.1
    optimized performance

  hm  14. mar. 2009 rev 1.2
    removed double assignments
*)
END_FUNCTION_BLOCK

(* ---- Measuring_Modules.ST ---- *)
(* @PATH := '\/Engineering\/measurements' *)
FUNCTION_BLOCK ALARM_2
(*
  ALARM_2 will check two pairs of limits and signal when the input is above or below a set limit.
  with the input HYS a hysteresis can be defined for all limits.

  version 1.1 11. mar. 2009
  programmer  hugo
  tested by   tobias
*)
  VAR_INPUT
    X : REAL;
    LO_1 : REAL;
    HI_1 : REAL;
    LO_2 : REAL;
    HI_2 : REAL;
    HYS : REAL;
  END_VAR
  VAR_OUTPUT
    Q1_LO : BOOL;
    Q1_HI : BOOL;
    Q2_LO : BOOL;
    Q2_HI : BOOL;
  END_VAR
  VAR
    tmp: REAL;
  END_VAR

  tmp := X - Hys * 0.5;
  IF tmp > LO_1 THEN Q1_LO := FALSE; END_IF;
  IF tmp > LO_2 THEN Q2_LO := FALSE; END_IF;
  IF tmp > HI_1 THEN Q1_HI := TRUE; END_IF;
  IF tmp > HI_2 THEN Q2_HI := TRUE; END_IF;
  tmp := tmp + hys;
  IF tmp < LO_1 THEN Q1_LO := TRUE; END_IF;
  IF tmp < LO_2 THEN Q2_LO := TRUE; END_IF;
  IF tmp < HI_1 THEN Q1_HI := FALSE; END_IF;
  IF tmp < HI_2 THEN Q2_HI := FALSE; END_IF;

(* revision history
  hm  19. may. 2008   rev 1.0
    original version

  hm  11. mar. 2009 rev 1.1
    improved code
*)
END_FUNCTION_BLOCK

(* @PATH := '\/Engineering\/measurements' *)
FUNCTION_BLOCK BAR_GRAPH
(*
  bar graph is a muti window comparator which displays an analog input signal on 8 digital outputs.
  only one output is active a any given time depending on the value of the input signal.
  the output can be of linear or logarithmic scale.

  version 1.2 6 jan 2008
  programmer  hugo
  tested by hans
*)
  VAR_INPUT
    X : REAL;
    rst : BOOL;
  END_VAR
  VAR_INPUT //???CONSTANT
    trigger_Low : REAL;
    trigger_High : REAL;
    Alarm_low : BOOL;
    Alarm_high : BOOL;
    log_scale : BOOL;
  END_VAR
  VAR_OUTPUT
    LOW, Q1, Q2, Q3, Q4, Q5, Q6, HIGH : BOOL;
    Alarm : BOOL;
    Status : BYTE;
  END_VAR
  VAR
    init : BOOL;
    T1, T2, T3, T4, T5 : REAL;
  END_VAR
  VAR_TEMP
    temp : REAL;
  END_VAR

  IF NOT init THEN
    init := TRUE;
    IF log_scale THEN
      temp := EXP(LN(Trigger_high / Trigger_low) * 0.166666666666666666666);
      T1 := trigger_low * temp;
      T2 := T1 * temp;
      T3 := T2 * temp;
      T4 := T3 * temp;
      T5 := T4 * temp;
    ELSE
      temp := (trigger_high - trigger_low) * 0.142857142;
      T1 := trigger_low + temp;
      T2 := T1 + temp;
      T3 := T2 + temp;
      T4 := T3 + temp;
      T5 := T4 + temp;
    END_IF;
  END_IF;

  (* clear outputs before checking *)
  Q1 := FALSE;
  Q2 := FALSE;
  Q3 := FALSE;
  Q4 := FALSE;
  Q5 := FALSE;
  Q6 := FALSE;
  status := 110;

  (* low, high and alarm can only be cleared with rst depending on alarm_low and alarm_high *)
  IF NOT alarm_low THEN low := FALSE; END_IF;
  IF NOT alarm_high THEN high := FALSE; END_IF;
  IF rst THEN
    alarm := FALSE;
    low := FALSE;
    high := FALSE;
  END_IF;

  (* check and set outputs *)
  IF X < trigger_low THEN
    Low := TRUE;
    status := 111;
    IF alarm_low THEN
      alarm := TRUE;
      status := 1;
    END_IF;
  ELSIF X < T1 THEN
    Q1 := TRUE;
  ELSIF x < t2 THEN
    Q2 := TRUE;
  ELSIF x < t3 THEN
    Q3 := TRUE;
  ELSIF x < T4 THEN
    Q4 := TRUE;
  ELSIF x < T5 THEN
    q5 := TRUE;
  ELSIF x < trigger_high THEN
    q6 := TRUE;
  ELSE
    high := TRUE;
    status := 112;
    IF alarm_high THEN
      alarm := TRUE;
      status := 2;
    END_IF;
  END_IF;

(* revision history
  hm  22. feb 2007  rev 1.0
    original version

  hm  2. dec 2007   rev 1.1
    chaged code for better performance

  hm  6. jan 2008   rev 1.2
    further performance improvement
*)
END_FUNCTION_BLOCK

(* @PATH := '\/Engineering\/measurements' *)
FUNCTION_BLOCK CALIBRATE
(*
  Calibrate allows for offset and scale calibration of an analog input.
  offset is calibrated to a stored reference Y_offset while CO is true.
  after the offset is calibrated, scale can be calibrated to a reference value Y_scale while CS is true.

  version 1.3 11. mar. 2009
  programmer  hugo
  tested by   hans
*)
  VAR_INPUT
    X : REAL;
    CO : BOOL;
    CS : BOOL;
  END_VAR
  VAR_INPUT //???CONSTANT
    Y_Offset : REAL;
    Y_Scale : REAL;
  END_VAR
  VAR_OUTPUT
    Y : REAL;
  END_VAR
  VAR_IN_OUT //???VAR RETAIN
    offset : REAL;
    Scale : REAL := 1.0;
  END_VAR

  (* check for calibration *)
  IF CO THEN
    OFFSET := Y_Offset - X;
  ELSIF CS THEN
    SCALE := Y_scale / (X + OFFSET);
  END_IF;
  (* calculate output *)
  Y := (X + OFFSET) * SCALE;

(* revision history
  hm 22.2.2007    rev 1.2
    changed VAR RETAIN PERSISTENT to VAR RETAIN for better compatibility
    wago lon contollers do not support persisitent

  hm  11. mar. 2009 rev 1.3
    changed real constants to use dot syntax
*)
END_FUNCTION_BLOCK

(* @PATH := '\/Engineering\/measurements' *)
FUNCTION_BLOCK CYCLE_TIME
(*
  this function block measures the cycle time and displays the last, min and max cycle time of the current task.
  the resolution is 1ms.
  the cycles output is a dword counter which counts the cycles.
  a rst pulse on the input will reset all data.

  version 1.2 16 sep 2007
  programmer  hugo
  tested by   hans
*)
  VAR_INPUT
    RST : BOOL;
  END_VAR
  VAR_OUTPUT
    ct_min : TIME;
    ct_max : TIME;
    ct_last : TIME;
    systime : TIME;
    sysdays : INT;
    cycles : DWORD;
  END_VAR
  VAR
    last_cycle : TIME;
    tx: TIME;
    init: BOOL;
  END_VAR

  tx := DWORD_TO_TIME(T_PLC_MS()) - last_cycle;
  IF rst THEN
    ct_min := t#10h;
    ct_max := t#0ms;
    cycles := 0;
  ELSIF last_cycle > t#0s THEN
    IF tx < ct_min THEN ct_min := tx;
    ELSIF tx > ct_max THEN ct_max := tx;
    END_IF;
    ct_last := tx;
  ELSIF ct_min = t#0s THEN
    ct_min := t#0s - t#1ms;
  END_IF;
  IF init THEN
    systime := systime + tx;
      IF systime >= t#1d THEN
        systime := systime - t#1d;
        sysdays := sysdays + 1;
      END_IF;
  END_IF;
  init := TRUE;
  last_cycle := last_cycle + tx;
  cycles := UDINT_TO_DWORD( DWORD_TO_UDINT(cycles) + 1);

(*  revision history
  hm 12.12.2006   rev 1.1
    added cycles output, a dword cycle counter.
  hm 10.3.2007      rev 1.2
    changed initialization of ct_min to t#10h for compatibility with siemens s7

  hm  16.9.2007   rev 1.2
    changed Time() in T_PLC_MS() for compatibility resons
*)
END_FUNCTION_BLOCK

(* @PATH := '\/Engineering\/measurements' *)
FUNCTION_BLOCK DT_SIMU
(*
  DT_SIMU simulates a real time clock and can be adjusted to different speeds
  it can also be used in simulation to simulate a real time clock.
  the peed of the clock can be increased or decreased to debug timers.
  with the input start a start date-time can be specified.

  version 1.2 8. mar. 2009
  programmer  hugo
  tested by   oscat
*)
  VAR_INPUT
    START : DT;
    SPEED : REAL := 1.0;
  END_VAR
  VAR_OUTPUT
    DTS : DT;
  END_VAR
  VAR
    tc : UDINT; //???DWORD;
    init: BOOL;
    last: UDINT; //???DWORD;
    tx: UDINT; //???DWORD;
    td: UDINT; //???DWORD;
  END_VAR

  (* read system timer *)
  tx := DWORD_TO_UDINT(T_PLC_MS());
  tc := REAL_TO_UDINT( UDINT_TO_REAL(tx - last) * speed);

  IF NOT init THEN
    init := TRUE;
    DTS := Start;
    tc := 0;
    last := tx;
  ELSIF SPEED = 0.0 THEN
    DTS := UDINT_TO_DT(DT_TO_UDINT(DTS) + 1);
  ELSIF tc >= 1000 THEN
    td := (tc / 1000) * 1000;
    DTS := ADD_DT_TIME( DTS, UDINT_TO_TIME(td));
    last := last + REAL_TO_UDINT( UDINT_TO_REAL(td) / speed);
  END_IF;

(* revision history
  hm  11. sep. 2008 rev 1.0
    original version

  hm  16. nov 2008  rev 1.1
    added type conversions for compatibility reasons

  hm  8.  mar. 2009 rev 1.2
    added increment by cycle mode
*)
END_FUNCTION_BLOCK

(* @PATH := '\/Engineering\/measurements' *)
FUNCTION_BLOCK FLOW_METER
(*
  Flow meter measures flow according to gated time or pulses.

  version 1.0 23. jan. 2011
  programmer  hugo
  tested by oscat
*)
  VAR_INPUT
    VX : REAL;
    E : BOOL;
    RST : BOOL;
  END_VAR
  VAR_INPUT //???CONSTANT
    PULSE_MODE : BOOL;
    UPDATE_TIME : TIME := t#1s;
  END_VAR
  VAR_OUTPUT
    F : REAL;
  END_VAR
  VAR_IN_OUT
    X : REAL;
    Y : UDINT;
  END_VAR
  VAR
    tx, tl : TIME;
    int1 : INTEGRATE;
    init: BOOL;
    e_last : BOOL;
    tmp: INT;
    x_last : REAL;
    y_last : UDINT;
  END_VAR

  IF NOT init THEN  (* init on power up *)
    init := TRUE;
    tl := tx;
    x_last := X;
    y_last := Y;
    int1.K := 2.7777777777777777E-4;
  END_IF;

  (* run integrator *)
  int1(E := NOT (RST OR PULSE_MODE) AND E, X := VX, Y := X);  (* gated operation *)

  IF RST THEN   (* reset *)
    X := 0.0;
    Y := 0;
    tl := tx;
    x_last := 0.0;
    y_last := 0;
  ELSIF E AND PULSE_MODE THEN (* check for pulse mode *)
    IF NOT e_last THEN X := X + VX; END_IF;
  END_IF;
  e_last := E;

  (* reduce X to be less than 1 and increase Y respectively *)
  IF X > 1.0 THEN
    tmp := FLOOR1(X);
    Y := Y + INT_TO_UDINT(tmp);
    X := X - INT_TO_REAL(tmp);
  END_IF;

  (* calculate the current flow *)
  tx := DWORD_TO_TIME(T_PLC_MS());
  IF tx - tl >= UPDATE_TIME AND UPDATE_TIME > t#0s THEN
    F := (UDINT_TO_REAL(Y - y_last) + X - x_last) / TIME_TO_REAL(tx - tl) * 3.6E6;
    y_last := Y;
    x_last := X;
    tl := tx;
  END_IF;

(* revision history
  hm  23. jan. 2011 rev 1.0
    original version
*)
END_FUNCTION_BLOCK

(* @PATH := '\/Engineering\/measurements' *)
FUNCTION_BLOCK M_D
(*
  m_d measures the time between a rising edge on start to a rising edge on stop and returs the last measured value on the output PT.
  a second output ET is starting from 0 at the rising edge of start and is counting up until the rising edge of stop occurs.
  the asynchronous input rst can reset the outputs at any time.
  tmax defines a timeout wich is the maximum measurable time between start and stop, if this time is exceeded the outputs will stay at 0.

  version 1.2 27. feb. 2009
  programmer  hugo
  tested by oscat
*)
  VAR_INPUT
    start : BOOL;
    stop : BOOL;
    tmax : TIME := t#10d;
    rst: BOOL;
  END_VAR
  VAR_OUTPUT
    PT : TIME;
    ET : TIME;
    run : BOOL;
  END_VAR
  VAR
    edge : BOOL;
    T0 : TIME;
    tx: TIME;
    startup: BOOL;
  END_VAR

  (* check for rst input *)
  IF rst OR et >= tmax THEN
    pt := t#0ms;
    et := t#0ms;
    startup := FALSE;
    run := FALSE;
  END_IF;

  (* avoid timers to start when input is true at startup *)
  IF NOT startup THEN
    edge := start;
    startup := TRUE;
  END_IF;

  (* read system timer *)
  tx := DWORD_TO_TIME(T_PLC_MS());

  (* detect rising edge on start *)
  IF start AND NOT edge AND NOT stop THEN
    t0 := tx;
    run := TRUE;
    pt := t#0s;
  ELSIF stop AND run THEN
    pt := et;
    run := FALSE;
  END_IF;
  edge := start;
  IF run THEN et := tx - t0; END_IF;

(* revision history
  hm    2.5.2007  rev 1.0
    original version

  hm    16.9.2007 rev 1.1
    changes time() to T_plc_ms() for compatibility reasons

  hm  27. feb 2009  rev 1.2
    deleted unnecessary init with 0
*)
END_FUNCTION_BLOCK

(* @PATH := '\/Engineering\/measurements' *)
FUNCTION_BLOCK M_T
(*
  m_t measures the with of a high pulse and returs the last measured pulse width on output PT.
  a second output ET is starting from 0 at the rising edge and counting up until the falling edge occurs and resetts et to 0.
  the asynchrtonous input rst can reset the outputs at any time.
  tmax defines a maximum measurable time, if this value is exceeded the outputs will be reset to 0.

  version 1.4 10. mar. 2009
  programmer  hugo
  tested by   oscat
*)
  VAR_INPUT
    IN : BOOL;
    TMAX : TIME := t#10d;
    RST : BOOL;
  END_VAR
  VAR_OUTPUT
    PT : TIME;
    ET: TIME;
  END_VAR
  VAR
    edge : BOOL;
    start : TIME;
    tx: TIME;
  END_VAR

  (* read system time *)
  tx := DWORD_TO_TIME(T_PLC_MS());

  IF RST OR ET >= TMAX THEN
    PT :=  t#0s;
    ET := t#0s;
  ELSIF IN THEN
    IF NOT edge THEN start := tx; END_IF;
    ET := tx - start;
  ELSE
    PT := ET;
  END_IF;
  edge := IN;

(* revision history
  hm  4. aug. 2006  rev 1.0
    original version

  hm  2. may. 2007  rev 1.1
    added init variable to avoid unreasonable measurement if falling edge occurs first.
    added et (elapsed time) output to count from 0 at rising edge until a falling edge resets et to 0.
    added reset input.

  hm  16. sep. 2007 rev 1.2
    changes time() to T_plc_ms() for compatibility reasons

  hm  17. dec. 2008 rev 1.3
    code optimized

  hm  10. mar. 2009 rev 1.4
    removed nested comments
    removed double assignments
*)
END_FUNCTION_BLOCK

(* @PATH := '\/Engineering\/measurements' *)
FUNCTION_BLOCK M_TX
(*
  this measures the timing of a signal
  TH is the high pulse width
  TL is the low pulse width
  DC is the duty cycle
  F is the frequency
  ET will start at 0 with a rising edge and count up till the next rising edge starts from 0 again.
  the acuracy depends on the cycle time of the sps and is limited to 1ms resolution.
  an asynchronous reset can reset all outputs to 0 at any time.
  the input tmax can configure a timeout for ET where the function block will outomatically reset itself.
  tmx is predefined to 10 days.

  version 1.4 11. mar. 2009
  programmer  oscat
  tested by   oscat
*)
  VAR_INPUT
    in: BOOL;
    tmax : TIME := t#10d;
    rst : BOOL;
  END_VAR
  VAR_OUTPUT
    TH : TIME;
    TL : TIME;
    DC : REAL;
    F: REAL;
    ET : TIME;
  END_VAR
  VAR
    edge : BOOL;
    start: TIME;
    stop:TIME;
    tx: TIME;
    rise : BOOL;
    fall : BOOL;
    startup: BOOL;
  END_VAR

  (* check FOR rst input *)
  IF rst OR (et >= tmax) THEN
    rise := FALSE;
    fall := FALSE;
    startup := FALSE;
    th := t#0ms;
    tl := t#0ms;
    DC := 0.0;
    F := 0.0;
    ET := t#0s;
  END_IF;

  (* avoid timers to start when input is true at startup *)
  IF NOT startup THEN
    edge := in;
    startup := TRUE;
  END_IF;

  (* read system timer *)
  tx := DWORD_TO_TIME(T_PLC_MS());

  (* edge trigger rising and falling edge *)
  IF in XOR edge THEN
    edge := in;
    (* rising edge starts measurement *)
    IF in THEN
      start := Tx;
      rise := TRUE;
      IF fall THEN tl := start - stop; END_IF;
      IF th > t#0ms AND tl > t#0ms THEN
        dc := TIME_TO_REAL(th) / TIME_TO_REAL(th+tl);
        f := 1000.0 / TIME_TO_REAL(th + tl);
      END_IF;
    (* falling edge starts second cycle measurement *)
    ELSE
      stop := Tx;
      fall := TRUE;
      IF rise THEN th := stop - start; END_IF;
      IF th > t#0ms AND tl > t#0ms THEN
        dc := TIME_TO_REAL(th) /  TIME_TO_REAL(th+tl);
        f := 1000.0 / TIME_TO_REAL(th + tl);
      END_IF;
    END_IF;
  END_IF;
  IF rise THEN et := tx - start; END_IF;

(* revision history
  hm  4. aug. 2006  rev 1.0
    original version

  hm  2. mai. 2007  rev 1.1
    made sure that no undefined values would be measured at startup conditions
    added output et
    added rst input
    added tmax input

  hm  16. sep. 2007 rev 1.2
    changes time() to T_plc_ms() for compatibility reasons

  hm  27. feb. 2009 rev 1.3
    deleted unnecessary init with 0

  hm  11. mar. 2009 rev 1.4
    changed real constants to use dot syntax
*)
END_FUNCTION_BLOCK

(* @PATH := '\/Engineering\/measurements' *)
FUNCTION_BLOCK METER
(*
  METER measures usage of power or similar values the output MX is the sum of the inputs over time.
  MX := sum over time of (I1 * P1 + I2 * P2)/D.
  a simple example is the consumption counter for a 2 stage oil burner where stage 1 is 10KW and stage 2 is 20KW.
  I1 and I2 decide which value is accounted for, I1 = True only counts P1, I2 is True counts P2
  and I1 and I2 is true counts P1 and P2.
  the meter can be used for all kind of consumption meters. P1 and P2 can change on the fly.

  version 1.4 8. mar. 2009
  programmer  oscat
  tested by oscat
*)
  VAR_INPUT
    M1, M2 : REAL;
    I1, I2 : BOOL;
    D : REAL := 1.0;
    RST : BOOL;
  END_VAR
  VAR_IN_OUT
    MX : REAL;
  END_VAR
  VAR
    MR : REAL2;
    MX1, MX2 : REAL; (* current consumption value on M1 and M2 *)
    tx: UDINT; //DWORD;
    last: UDINT; //DWORD;
    tc: REAL;
    init: BOOL;
  END_VAR

  (* measure the last cycle time and make sure we onle execute once every millisecond *)
  tx := DWORD_TO_UDINT( T_PLC_MS());
  IF NOT init THEN
    init := TRUE;
    last := tx;
    mr.RX := mx;
    mr.R1 := 0.0;
  ELSIF tx = last THEN
    RETURN;
  ELSE
    tc := UDINT_TO_REAL(tx - last) * 0.001;
  END_IF;
  last := tx;

  (* reset *)
  IF rst THEN
    mr.R1 := 0.0;
    mr.RX := 0.0;
  ELSE
    (* current consumption measurement *)
    IF I1 THEN MX1 := M1; ELSE MX1 := 0.0; END_IF;
    IF I2 THEN MX2 := M2; ELSE MX2 := 0.0; END_IF;
    (* add up the current values in a double real *)
    MR := R2_ADD(MR,(SEL(I1,0.0,mx1) + SEL(I2, 0.0, mx2)) / D * TC);
    (* set the current output value *)
    MX := mr.RX;
  END_IF;

(* revision history
  hm  16. sep.2007    rev 1.0
    original version

  hm  7. feb 2008   rev 1.1
    use new version of ft_int to avoid a counting stop at high values
    deleted unnecessary limits

  hm  24. mar. 2008 rev 1.2
    use data_type real2 to extend accuracy to 15 digits total
    do not use ft_int which adds unnecessary overhead

  hm  8. feb. 2009  rev 1.3
    changed mx to be I/O
    make sure calculation works for cycle times < 1 ms

  hm  8. mar. 2009  rev 1.4
    last was not updated
    code improvements
*)
END_FUNCTION_BLOCK

(* @PATH := '\/Engineering\/measurements' *)
FUNCTION_BLOCK METER_STAT
(*
  METER_STAT runs statistics of a metered value, it calculates the current week, day, month and year consumption and stores the corresponding last day, week, month and year value.

  version 1.3 18. jul. 2009
  programmer  oscat
  tested by   oscat
*)
  VAR_INPUT
    IN : REAL;
    DI : DATE;
    RST : BOOL;
  END_VAR
  VAR_IN_OUT
    Last_Day : REAL;
    Current_Day : REAL;
    Last_Week : REAL;
    Current_Week : REAL;
    Last_Month : REAL;
    Current_Month : REAL;
    Last_Year : REAL;
    Current_Year : REAL;
  END_VAR
  VAR_IN_OUT //!!!VAR RETAIN
    Year_Start : REAL;
    Month_Start : REAL;
    Week_Start : REAL;
    Day_Start : REAL;
    last_run: DATE;
  END_VAR

  IF rst THEN
    Last_Day := 0.0;
    Current_Day := 0.0;
    Day_start := IN;
    Last_week := 0.0;
    Current_week := 0.0;
    Week_start := in;
    Last_month := 0.0;
    Current_month := 0.0;
    month_start := in;
    last_year := 0.0;
    current_year := 0.0;
    year_start := in;
  ELSE
    Current_Day := IN - Day_Start;
    Current_Week := In - Week_Start;
    Current_Month := IN - Month_Start;
    Current_Year := IN - Year_Start;
  END_IF;

  IF YEAR_OF_DATE1(DI) > YEAR_OF_DATE1(last_run) THEN
    (* a new year has started *)
    last_year := current_year;
    current_year := 0.0;
    year_start := in;
    last_month := current_month;
    current_month := 0.0;
    month_start := in;
    last_day := current_day;
    current_day := 0.0;
    day_start := in;
  ELSIF MONTH_OF_DATE1(DI) > MONTH_OF_DATE1(last_run) THEN
    (* a new month has started, january is alrerady done by year change *)
    last_month := current_month;
    current_month := 0.0;
    month_start := in;
    last_day := current_day;
    current_day := 0.0;
    day_start := in;
  ELSIF DAY_OF_YEAR1(di) > DAY_OF_YEAR1(last_run) THEN
    (* day has chaged, first day of year and first day of month has already been taken care of *)
    last_day := current_day;
    current_day := 0.0;
    day_start := in;
  END_IF;
  IF DAY_OF_WEEK1(DI) < DAY_OF_WEEK1(last_run) THEN
    (* a new week has started *)
    last_week := current_week;
    current_week := 0.0;
    week_start := in;
  END_IF;
  last_run := di;

(* revision history
  hm  16. sep. 2007 rev 1.0
    original version

  hm  7. oct. 2008  rev 1.1
    changed function year_to_year_of_date
    changed function month to month_of_date
    changed function weekday to day_of_week

  hm  11. mar. 2009 rev 1.2
    changed real constants to use dot syntax

  hm  18. jul. 2009 rev 1.3
    changes all outputs to be I/O
*)
END_FUNCTION_BLOCK

(* @PATH := '\/Engineering\/measurements' *)
FUNCTION_BLOCK ONTIME
(*
  ONTIME measures the ontime of a signal in seconds.
  the output SECONDS is of type DWORD which results in a total measurement range of 1 second up to 136 years.
  internally ontime works with a resolution of milliseconds

  version 2.5 18. mar. 2011
  programmer  oscat
  tested by   tobias
*)
  VAR_INPUT
    IN : BOOL;
    RST : BOOL;
  END_VAR
  VAR_IN_OUT
    SECONDS : UDINT;
    CYCLES : UDINT;
  END_VAR
  VAR
    tx: UDINT; //DWORD;
    last : UDINT; //DWORD;
    edge : BOOL;
    init: BOOL;
    ms: UDINT; //DWORD;
  END_VAR

  (* read system time *)
  tx := DWORD_TO_UDINT( T_PLC_MS());

  (* make sure the first cycle works correctly *)
  IF NOT init THEN
    init := TRUE;
    last := tx;
    ms := 0;
  END_IF;
  IF RST THEN
    SECONDS := 0;
    CYCLES := 0;
    last := tx;
    ms := 0;
  ELSIF IN THEN
    (* add the current milliseconds *)
    ms := (tx - last) + ms;
    IF ms >= 1000 THEN
      seconds := seconds + 1;
      ms := ms - 1000;
    END_IF;
    cycles := cycles + BOOL_TO_UDINT(NOT edge);
  END_IF;
  last := tx;
  edge := in;

(* revision history
  hm 22.2.2007    rev 1.1
    changed VAR RETAIN PERSISTENT to VAR RETAIN for better compatibility
    wago lon contollers do not support persisitent

  hm 2.8.2007   rev 1.2
    adding time up in a real number will automatically lead to the point where
    small time scales like the cycle time will be below the resolution of real and therefore
    ontime would not increase in small steps as necessary
    the time is now measured internally in two  dwords and be converted to real only for
    output purposes.
    deleted the variable power because it was unnecessary

  hm  16.9.2007   rev 1.3
    changes time() to T_plc_ms() for compatibility reasons

  hm  2. dec. 2007  rev 1.4
    chaged code for better performance

  hm  16. mar. 2008 rev 1.5
    added type conversions to avoid warnings under codesys 3.0

  hm  21. oct. 2008 rev 2.0
    changed module for much better performance and allow for external result storage

  hm  10. nov. 2008 rev 2.1
    increased internal resolution to milliseconds

  hm  16. nov. 2008 rev 2.2
    changed typecast to avoid warnings

  hm  17. dec. 2008 rev 2.3
    fixed an error when in would be true for more then 49 days

  hm  17. jan 2011  rev 2.4
    init will not clear seconds and cycles, only rst clears these values

  hm  18. mar. 2011 rev 2.5
    reset was not working
*)
END_FUNCTION_BLOCK

(* @PATH := '\/Engineering\/measurements' *)
FUNCTION_BLOCK TC_MS
(*
  TC_MS delivers the time it was last called on the output TC in Milliseconds.

  version 1.0 13 mar 2008
  programmer  hugo
  tested by   tobias
*)
  VAR_OUTPUT
    TC : DWORD;
  END_VAR
  VAR
    init: BOOL;
    tx: UDINT; //DWORD;
    last: UDINT; //DWORD;
  END_VAR

  (* read system timer *)
  tx := DWORD_TO_UDINT( T_PLC_MS());

  IF NOT init THEN
    init := TRUE;
    TC := 0;
  ELSE
    tc := UDINT_TO_DWORD(tx - last);
  END_IF;
  last := tx;

(* revision history
  hm    13. mar. 2008 rev 1.0
    original version
*)
END_FUNCTION_BLOCK

(* @PATH := '\/Engineering\/measurements' *)
FUNCTION_BLOCK TC_S
(*
  TC_S delivers the time it was last called on the output TC in seconds.

  version 1.2 11. mar. 2009
  programmer  hugo
  tested by   tobias
*)
  VAR_OUTPUT
    TC : REAL;
  END_VAR
  VAR
    init: BOOL;
    tx: UDINT; //DWORD;
    last: UDINT; //DWORD;
  END_VAR

  (* read system timer *)
  tx := DWORD_TO_UDINT( T_PLC_US());

  IF NOT init THEN
    init := TRUE;
    TC := 0.0;
  ELSE
    tc := UDINT_TO_REAL(tx - last)*1.0E-6;
  END_IF;
  last := tx;

(* revision history
  hm  13. mar. 2008 rev 1.0
    original version

  hm  16. mar 2008  rev 1.1
    added type conversion to avoid warnings under codesys 3.0

  hm  11. mar. 2009 rev 1.2
    changed real constants to use dot syntax
*)
END_FUNCTION_BLOCK

(* @PATH := '\/Engineering\/measurements' *)
FUNCTION_BLOCK TC_US
(*
  TC_US delivers the time it was last called on the output TC in Microseconds.

  version 1.0 13 mar 2008
  programmer  hugo
  tested by   tobias
*)
  VAR_OUTPUT
    TC : DWORD;
  END_VAR
  VAR
    init: BOOL;
    tx: UDINT; //DWORD;
    last: UDINT; //DWORD;
  END_VAR

  (* read system timer *)
  tx := DWORD_TO_UDINT( T_PLC_US());

  IF NOT init THEN
    init := TRUE;
    TC := 0;
  ELSE
    tc := UDINT_TO_DWORD(tx - last);
  END_IF;
  last := tx;

(* revision history
  hm    13. mar. 2008 rev 1.0
    original version
*)
END_FUNCTION_BLOCK

(* ---- Memory_Modules.ST ---- *)
(* @PATH := '\/Logic\/memory' *)
FUNCTION_BLOCK FIFO_16
(*
  16 Dword FIFO memory

  version 2.0 24. jul. 2009
  programmer  hugo
  tested by   oscat
*)
  VAR_INPUT
    Din : DWORD;
    E : BOOL := TRUE;
    RD : BOOL;
    WD : BOOL;
    RST : BOOL;
  END_VAR
  VAR_OUTPUT
    Dout : DWORD;
    EMPTY : BOOL := TRUE;
    FULL : BOOL;
  END_VAR
  VAR CONSTANT
    n : INT := 16;  (* changing this value will chage the number of stored elements in the fifo *)
  END_VAR
  VAR
    fifo : ARRAY[0..n] OF DWORD;
    pr : INT;
    pw : INT;
  END_VAR

  IF RST THEN
    pw := pr;
    FULL := FALSE;
    EMPTY := TRUE;
    Dout := 0;
  ELSIF E THEN
    IF NOT EMPTY AND RD THEN
      Dout := fifo[pr];
      pr := INC1(pr,n);
      EMPTY := pr = pw;
      FULL := FALSE;
    END_IF;
    IF NOT FULL AND WD THEN
      fifo[pw] := Din;
      pw := INC1(pw,n);
      FULL := pw = pr;
      EMPTY := FALSE;
    END_IF;
  END_IF;

(* revision history
  hm  4. aug. 2006  rev 1.0
    original version

  hm  19. feb 2008  rev 1.1
    performance improvements

  hm  17. oct. 2008 rev 1.2
    improved performance

  ks  27. oct. 2008 rev 1.3
    optimized coding

  hm  14. mar. 2009 rev 1.4
    removed double assignments

  hm 24. jul. 2009  rev 2.0
    chaged inputs E and WR to E, WD and WR
    allow read and write in one cycle
*)
END_FUNCTION_BLOCK

(* @PATH := '\/Logic\/memory' *)
FUNCTION_BLOCK FIFO_32
(*
  32 Dword FIFO memory

  version 2.0 24. jul. 2009
  programmer  hugo
  tested by   oscat
*)
  VAR_INPUT
    Din : DWORD;
    E : BOOL := TRUE;
    RD : BOOL;
    WD : BOOL;
    RST : BOOL;
  END_VAR
  VAR_OUTPUT
    Dout : DWORD;
    EMPTY : BOOL := TRUE;
    FULL : BOOL;
  END_VAR
  VAR CONSTANT
    n : INT := 32;  (* changing this value will chage the number of stored elements in the fifo *)
  END_VAR
  VAR
    fifo : ARRAY[0..n] OF DWORD;
    pr : INT;
    pw : INT;
  END_VAR

  IF RST THEN
    pw := pr;
    FULL := FALSE;
    EMPTY := TRUE;
    Dout := 0;
  ELSIF E THEN
    IF NOT EMPTY AND RD THEN
      Dout := fifo[pr];
      pr := INC1(pr,n);
      EMPTY := pr = pw;
      FULL := FALSE;
    END_IF;
    IF NOT FULL AND WD THEN
      fifo[pw] := Din;
      pw := INC1(pw,n);
      FULL := pw = pr;
      EMPTY := FALSE;
    END_IF;
  END_IF;

(* revision history
  hm  4. aug. 2006  rev 1.0
    original version

  hm  19. feb 2008  rev 1.1
    performance improvements

  hm  17. oct. 2008 rev 1.2
    improved performance

  ks  27. oct. 2008 rev 1.3
    improved code

  hm  14. mar. 2009 rev 1.4
    removed double assignments

  hm 24. jul. 2009  rev 2.0
    chaged inputs E and WR to E, WD and WR
    allow read and write in one cycle
*)
END_FUNCTION_BLOCK

(* @PATH := '\/Logic\/memory' *)
FUNCTION_BLOCK STACK_16
(*
  16 Dword STACK memory

  version 2.0 25. jul 2009
  programmer  hugo
  tested by   oscat
*)
  VAR_INPUT
    Din : DWORD;
    E : BOOL := TRUE;
    RD : BOOL;
    WD : BOOL;
    RST : BOOL;
  END_VAR
  VAR_OUTPUT
    Dout : DWORD;
    EMPTY : BOOL := TRUE;
    FULL : BOOL;
  END_VAR
  VAR CONSTANT
    n : INT := 15;  (* changing this value will chage the number of stored elements in the fifo *)
  END_VAR
  VAR
    stack : ARRAY[0..n] OF DWORD;
    pt : INT;
  END_VAR

  IF RST THEN
    (* asynchronous reset for the fifo *)
    pt := 0;
    EMPTY := TRUE;
    FULL := FALSE;
    Dout := 0;
  ELSIF E THEN
    IF NOT EMPTY AND RD THEN
      (* read one element *)
      pt := pt - 1;
      Dout := stack[pt];
      EMPTY := pt = 0;
      FULL := FALSE;
    END_IF;
    IF NOT FULL AND WD THEN
      (* write one element *)
      stack[pt] := Din;
      pt := pt + 1;
      FULL := pt > n;
      EMPTY := FALSE;
    END_IF;
  END_IF;

(* revision history
  hm  4. aug. 2006  rev 1.0
    original version

  hm  19. feb 2008  rev 1.1
    performance improvements

  hm  17. oct. 2008 rev 1.2
    deleted unnecessary init with 0

  hm  27. oct. 2008 rev 1.3
    optimized performance

  hm  25. jul 2009  rev 2.0
    changed inputs to allow simultsaneous read and write
*)
END_FUNCTION_BLOCK

(* @PATH := '\/Logic\/memory' *)
FUNCTION_BLOCK STACK_32
(*
  32 Dword STACK memory

  version 2.0 25. jul 2009
  programmer  hugo
  tested by   oscat
*)
  VAR_INPUT
    Din : DWORD;
    E : BOOL := TRUE;
    RD : BOOL;
    WD : BOOL;
    RST : BOOL;
  END_VAR
  VAR_OUTPUT
    Dout : DWORD;
    EMPTY : BOOL := TRUE;
    FULL : BOOL;
  END_VAR
  VAR CONSTANT
    n : INT := 31;  (* changing this value will chage the number of stored elements in the fifo *)
  END_VAR
  VAR
    stack : ARRAY[0..n] OF DWORD;
    pt : INT;
  END_VAR

  IF RST THEN
    (* asynchronous reset for the fifo *)
    pt := 0;
    EMPTY := TRUE;
    FULL := FALSE;
    Dout := 0;
  ELSIF E THEN
    IF NOT EMPTY AND RD THEN
      (* read one element *)
      pt := pt - 1;
      Dout := stack[pt];
      EMPTY := pt = 0;
      FULL := FALSE;
    END_IF;
    IF NOT FULL AND WD THEN
      (* write one element *)
      stack[pt] := Din;
      pt := pt + 1;
      FULL := pt > n;
      EMPTY := FALSE;
    END_IF;
  END_IF;

(* revision history
  hm  4. aug. 2006  rev 1.0
    original version

  hm  19. feb 2008  rev 1.1
    performance improvements

  hm  17. oct. 2008 rev 1.2
    deleted unnecessary init with 0

  ks  27. oct. 2008 rev 1.3
    optimized performance

  hm  25. jul 2009  rev 2.0
    changed inputs to allow simultsaneous read and write
*)
END_FUNCTION_BLOCK

(* ---- Other_Functions.ST ---- *)
TYPE
  OSCAT_BASIC_ARRAY0_3_OF_esr_data : ARRAY [0..3] OF esr_data;
END_TYPE

(* @PATH := '\/Other' *)
FUNCTION_BLOCK ESR_COLLECT
(*
  ESR_collect collects esr data from up to 8 esr_mon modules and stroes them in an output array.
  the output pos will display the position of the last element in the array. if the array is empty, pos = -1
  when to buffer is read by followon modules. pos has to be reset to -1
  if the array will be full, the buffer will be refilled starting at position 0.

  version 1.4 1. dec. 2009
  programmer  hugo
  tested by   tobias
*)
  VAR_INPUT
    ESR_0, ESR_1, ESR_2, ESR_3, ESR_4, ESR_5, ESR_6, ESR_7 : ARRAY [0..3] OF esr_data;
    rst : BOOL;
  END_VAR
  VAR_IN_OUT
    pos : INT;
  END_VAR
  VAR_OUTPUT
    ESR_OUT : ARRAY[0..31] OF esr_data;
  END_VAR
  VAR CONSTANT
    max_in : INT := 3; (* max limit of input array *)
    max_out : INT := 32; (* number of elements in array *)
  END_VAR
  VAR
    cnt : INT := -1;
  END_VAR

  IF rst OR cnt < 0 THEN
    pos := -1;
  ELSE
    FOR cnt := 0 TO max_in DO
    IF esr_0[cnt].typ > 0 THEN pos := INC1(pos, max_out); esr_out[pos] := esr_0[cnt]; END_IF;
    IF esr_1[cnt].typ > 0 THEN pos := INC1(pos, max_out); esr_out[pos] := esr_1[cnt]; END_IF;
    IF esr_2[cnt].typ > 0 THEN pos := INC1(pos, max_out); esr_out[pos] := esr_2[cnt]; END_IF;
    IF esr_3[cnt].typ > 0 THEN pos := INC1(pos, max_out); esr_out[pos] := esr_3[cnt]; END_IF;
    IF esr_4[cnt].typ > 0 THEN pos := INC1(pos, max_out); esr_out[pos] := esr_4[cnt]; END_IF;
    IF esr_5[cnt].typ > 0 THEN pos := INC1(pos, max_out); esr_out[pos] := esr_5[cnt]; END_IF;
    IF esr_6[cnt].typ > 0 THEN pos := INC1(pos, max_out); esr_out[pos] := esr_6[cnt]; END_IF;
    IF esr_7[cnt].typ > 0 THEN pos := INC1(pos, max_out); esr_out[pos] := esr_7[cnt]; END_IF;
     END_FOR;
  END_IF;

(* revision history
  hm  26.jan 2007 rev 1.0
    original version

  hm  8. dec 2007 rev 1.1
    added reset input

  ks  27. oct. 2008 rev 1.2
    optimized code for performance

  ks  12. nov. 2009 rev 1.3
    output pos was not pointing to last value

  hm  1. dec. 2009  rev 1.4
    changed pos to be I/O
    reduced output array size to 32 elements
*)
END_FUNCTION_BLOCK

(* @PATH := '\/Other' *)
FUNCTION_BLOCK ESR_MON_B8
(*
  ESR_mon_B8 monitores up to 8 binary inputs and reports changes with time stamd and adress label.
  the module checks 8 inputs for a change and reports all changes with time and adress stamp to the output.
  4 events maximum can be collected at once within the same cycle

  version 1.3 1. dec. 2009
  programmer  hugo
  tested by   tobias
*)
  VAR_INPUT
    s0, s1, s2, s3, s4, s5, s6, s7 : BOOL;
    DT_in : DT;
  END_VAR
  VAR_INPUT //???CONSTANT
    a0, a1, a2, a3, a4, a5, a6, a7 : STRING[10];
  END_VAR
  VAR_OUTPUT
    ESR_Flag : BOOL;
  END_VAR
  VAR_IN_OUT
    ESR_Out: OSCAT_BASIC_ARRAY0_3_OF_esr_data; // ARRAY [0..3] OF esr_data;
  END_VAR
  VAR
    x0, x1, x2, x3, x4, x5, x6, x7 : BOOL;
    tx: TIME;
    cnt : INT;
  END_VAR

  (* read system timer *)
  tx := DWORD_TO_TIME(T_PLC_MS());

  ESR_Flag := FALSE;
  esr_out[3].typ := 0;
  esr_out[2].typ := 0;
  esr_out[1].typ := 0;
  esr_out[0].typ := 0;
  cnt := 0;

  (* check if inputs have chaged and fill buffer *)
  IF s0 <> X0 THEN
    esr_out[cnt].typ := USINT_TO_BYTE(10 + BOOL_TO_USINT(s0));
    esr_out[cnt].adress := a0;
    esr_out[cnt].DS := DT_in;
    esr_out[cnt].TS := TX;
    X0 := S0;
    cnt := cnt + 1;
    esr_flag := TRUE;
  END_IF;
  IF s1 <> X1 THEN
    esr_out[cnt].typ := USINT_TO_BYTE(10 + BOOL_TO_USINT(s1));
    esr_out[cnt].adress := a1;
    esr_out[cnt].DS := DT_in;
    esr_out[cnt].TS := TX;
    X1 := S1;
    cnt := cnt + 1;
    esr_flag := TRUE;
  END_IF;
  IF s2 <> X2 THEN
    esr_out[cnt].typ := USINT_TO_BYTE(10 + BOOL_TO_USINT(s2));
    esr_out[cnt].adress := a2;
    esr_out[cnt].DS := DT_in;
    esr_out[cnt].TS := TX;
    X2 := S2;
    cnt := cnt + 1;
    esr_flag := TRUE;
  END_IF;
  IF s3 <> X3 THEN
    esr_out[cnt].typ := USINT_TO_BYTE(10 + BOOL_TO_USINT(s3));
    esr_out[cnt].adress := a3;
    esr_out[cnt].DS := DT_in;
    esr_out[cnt].TS := TX;
    X3 := S3;
    cnt := cnt + 1;
    esr_flag := TRUE;
  END_IF;
  IF s4 <> X4 AND cnt < 4 THEN
    esr_out[cnt].typ := USINT_TO_BYTE(10 + BOOL_TO_USINT(s4));
    esr_out[cnt].adress := a4;
    esr_out[cnt].DS := DT_in;
    esr_out[cnt].TS := TX;
    X4 := S4;
    cnt := cnt + 1;
    esr_flag := TRUE;
  END_IF;
  IF s5 <> X5  AND cnt < 4 THEN
    esr_out[cnt].typ := USINT_TO_BYTE(10 + BOOL_TO_USINT(s5));
    esr_out[cnt].adress := a5;
    esr_out[cnt].DS := DT_in;
    esr_out[cnt].TS := TX;
    X5 := S5;
    cnt := cnt + 1;
    esr_flag := TRUE;
  END_IF;
  IF s6 <> X6  AND cnt < 4 THEN
    esr_out[cnt].typ := USINT_TO_BYTE(10 + BOOL_TO_USINT(s6));
    esr_out[cnt].adress := a6;
    esr_out[cnt].DS := DT_in;
    esr_out[cnt].TS := TX;
    X6 := S6;
    cnt := cnt + 1;
    esr_flag := TRUE;
  END_IF;
  IF s7 <> X7  AND cnt < 4 THEN
    esr_out[cnt].typ := USINT_TO_BYTE(10 + BOOL_TO_USINT(s7));
    esr_out[cnt].adress := a7;
    esr_out[cnt].DS := DT_in;
    esr_out[cnt].TS := TX;
    X7 := S7;
    cnt := cnt + 1;
    esr_flag := TRUE;
  END_IF;

(* revision history
  hm  26. jan 2007  rev 1.0
    original version

  hm  17. sep 2007  rev 1.1
    replaced time() with T_PLC_MS() for compatibility reasons

  hm  22. oct. 2008 rev 1.2
    optimized code

  hm  1.dec. 2009 rev 1.3
    changed esr_out to be I/O
*)
END_FUNCTION_BLOCK

(* @PATH := '\/Other' *)
FUNCTION_BLOCK ESR_MON_R4
(*
  ESR_mon_R4 monitores up to 4 Real inputs and reports changes with time stamd and adress label.
  the module checks 4 inputs for a change of more than the specified sensitivity S and reports all changes with time and adress stamp to the output.

  version 1.4 1. dec. 2009
  programmer  hugo
  tested by   tobias
*)
  VAR_INPUT
    R0, R1, R2, R3 : REAL;
    DT_in : DT;
  END_VAR
  VAR_INPUT //???CONSTANT
    a0, a1, a2, a3 : STRING[10];
    s0, s1, s2, s3 : REAL;
  END_VAR
  VAR_OUTPUT
    ESR_Flag : BOOL;
  END_VAR
  VAR_IN_OUT
    ESR_Out: OSCAT_BASIC_ARRAY0_3_OF_esr_data; // ARRAY [0..3] OF esr_data;
  END_VAR
  VAR
    p0, p1, p2, p3 : PTR_TO DWORD;
    x0, x1, x2, x3 : REAL;
    tx: TIME;
    cnt : INT;
  END_VAR

  (* read system timer *)
  tx := DWORD_TO_TIME(T_PLC_MS());
  P0 := ADR(R0);
  P1 := ADR(R1);
  P2 := ADR(R2);
  P3 := ADR(R3);

  ESR_Flag := FALSE;
  esr_out[3].typ := 0;
  esr_out[2].typ := 0;
  esr_out[1].typ := 0;
  esr_out[0].typ := 0;
  cnt := 0;

  (* check if inputs have chaged and fill buffer *)
  IF DIFFER(R0,  X0, S0) THEN
    esr_out[cnt].typ := 20;
    esr_out[cnt].adress := a0;
    esr_out[cnt].DS := DT_in;
    esr_out[cnt].TS := TX;
    esr_out[cnt].data[0] := Byte_of_Dword(P0^,0);
    esr_out[cnt].data[1] := Byte_of_Dword(P0^,1);
    esr_out[cnt].data[2] := Byte_of_Dword(P0^,2);
    esr_out[cnt].data[3] := Byte_of_Dword(P0^,3);
    X0 := R0;
    cnt := cnt + 1;
    esr_flag := TRUE;
  END_IF;
  IF differ(R1,  X1, S1) THEN
    esr_out[cnt].typ := 20;
    esr_out[cnt].adress := a1;
    esr_out[cnt].DS := DT_in;
    esr_out[cnt].TS := TX;
    esr_out[cnt].data[0] := Byte_of_Dword(P1^,0);
    esr_out[cnt].data[1] := Byte_of_Dword(P1^,1);
    esr_out[cnt].data[2] := Byte_of_Dword(P1^,2);
    esr_out[cnt].data[3] := Byte_of_Dword(P1^,3);
    X1 := R1;
    cnt := cnt + 1;
    esr_flag := TRUE;
  END_IF;
  IF differ(R2,  X2, S2) THEN
    esr_out[cnt].typ := 20;
    esr_out[cnt].adress := a2;
    esr_out[cnt].DS := DT_in;
    esr_out[cnt].TS := TX;
    esr_out[cnt].data[0] := Byte_of_Dword(P2^,0);
    esr_out[cnt].data[1] := Byte_of_Dword(P2^,1);
    esr_out[cnt].data[2] := Byte_of_Dword(P2^,2);
    esr_out[cnt].data[3] := Byte_of_Dword(P2^,3);
    X2 := R2;
    cnt := cnt + 1;
    esr_flag := TRUE;
  END_IF;
  IF DIFFER(R3,  X3, S3) THEN
    esr_out[cnt].typ := 20;
    esr_out[cnt].adress := a3;
    esr_out[cnt].DS := DT_in;
    esr_out[cnt].TS := TX;
    esr_out[cnt].data[0] := Byte_of_Dword(P3^,0);
    esr_out[cnt].data[1] := Byte_of_Dword(P3^,1);
    esr_out[cnt].data[2] := Byte_of_Dword(P3^,2);
    esr_out[cnt].data[3] := Byte_of_Dword(P3^,3);
    X3 := R3;
    cnt := cnt + 1;
    esr_flag := TRUE;
  END_IF;

(* revision history
  hm  26. jan 2007  rev 1.0
    original version

  hm  17. sep. 2007   rev 1.1
    replaced time() with T_PLC_MS() for compatibility reasons

  hm  8. dec. 2007    rev 1.2
    corrected an error while esr typ would not be set

  hm  16. mar. 2008   rev 1.3
    deleted wrong conversion real_to_dword

  hm  1. dec 2009   rev 1.4
    changed esr_out to be I/O
*)
END_FUNCTION_BLOCK

(* @PATH := '\/Other' *)
FUNCTION STATUS_TO_ESR : esr_data
(*
  status_to_esr creates esr data from a status byte.

  version 1.0 6 oct 2006
  programmer  hugo
  tested by   tobias
*)
  VAR_INPUT
    status : BYTE;
    adress : STRING[10];
    DT_in : DT;
    TS : TIME;
  END_VAR

  IF status < 100 THEN
    status_to_ESR.typ := 1;
  ELSIF status < 200 THEN
    status_to_ESR.typ := 2;
  ELSE
    status_to_ESR.typ := 3;
  END_IF;
  status_to_ESR.adress:= adress;
  status_to_ESR.DS := DT_in;
  status_to_ESR.TS := TS;
  status_to_ESR.data[0] := status;

END_FUNCTION

(* @PATH := '\/Other' *)
FUNCTION_BLOCK ESR_MON_X8
(*
  ESR_MON_X8 is a status and error collector.
  the module checks 8 status inputs for a change and reports up to 4 input changes with time and adress stamp to the output.
  the mode can be
  1 for error only
  2 for error and status
  3 for error, status and debug
  the adress label of the 8 inputs can be configured individually.

  version 1.2 1. dec. 2009
  programmer  hugo
  tested by   tobias
*)
  VAR_INPUT
    s0, s1, s2, s3, s4, s5, s6, s7 : BYTE;
    DT_in : DT;
    Mode : BYTE := 3;
  END_VAR
  VAR_INPUT //???CONSTANT
    a0, a1, a2, a3, a4, a5, a6, a7 : STRING[10];
  END_VAR
  VAR_OUTPUT
    ESR_Flag : BOOL;
  END_VAR
  VAR_IN_OUT
    ESR_Out: OSCAT_BASIC_ARRAY0_3_OF_esr_data; // ARRAY [0..3] OF esr_data;
  END_VAR
  VAR
    x0, x1, x2, x3, x4, x5, x6, x7 : BYTE;
    tx: TIME;
    cnt : INT;
  END_VAR

  (* read system timer *)
  tx := DWORD_TO_TIME(T_PLC_MS());

  ESR_Flag := FALSE;
  esr_out[3].typ := 0;
  esr_out[2].typ := 0;
  esr_out[1].typ := 0;
  esr_out[0].typ := 0;
  cnt := 0;

  (* check if inputs have chaged and fill buffer *)
  IF (s0 <> X0) AND ((s0 < 100) OR ((S0 > 99) AND (S0 < 200) AND (mode >= 2)) OR ((S0 > 199) AND (mode = 3))) THEN
    esr_out[cnt] := status_to_ESR(s0, a0, DT_in, TX);
    X0 := S0;
    cnt := cnt + 1;
    esr_flag := TRUE;
  END_IF;
  IF (s1 <> X1) AND ((s1 < 100) OR ((S1 > 99) AND (S1 < 200) AND (mode >= 2)) OR ((S1 > 199) AND (mode = 3))) THEN
    esr_out[cnt] := status_to_ESR(s1, a1, DT_in, TX);
    X1 := S1;
    cnt := cnt + 1;
    esr_flag := TRUE;
  END_IF;
  IF (s2 <> X2) AND ((s2 < 100) OR ((S2 > 99) AND (S2 < 200) AND (mode >= 2)) OR ((S2 > 199) AND (mode = 3))) THEN
    esr_out[cnt] := status_to_ESR(s2, a2, DT_in, TX);
    X2 := S2;
    cnt := cnt + 1;
    esr_flag := TRUE;
  END_IF;
  IF (s3 <> X3) AND ((s3 < 100) OR ((S3 > 99) AND (S3 < 200) AND (mode >= 2)) OR ((S3 > 199) AND (mode = 3))) THEN
    esr_out[cnt] := status_to_ESR(s3, a3, DT_in, TX);
    X3 := S3;
    cnt := cnt + 1;
    esr_flag := TRUE;
  END_IF;
  IF (cnt < 4) AND (s4 <> X4) AND ((s4 < 100) OR ((S4 > 99) AND (S4 < 200) AND (mode >= 2)) OR ((S4 > 199) AND (mode = 3))) THEN
    esr_out[cnt] := status_to_ESR(s4, a4, DT_in, TX);
    X4 := S4;
    cnt := cnt + 1;
    esr_flag := TRUE;
  END_IF;
  IF (cnt < 4) AND (s5 <> X5) AND ((s5 < 100) OR ((S5 > 99) AND (S5 < 200) AND (mode >= 2)) OR ((S5 > 199) AND (mode = 3))) THEN
    esr_out[cnt] := status_to_ESR(s5, a5, DT_in, TX);
    X5 := S5;
    cnt := cnt + 1;
    esr_flag := TRUE;
  END_IF;
  IF (cnt < 4) AND (s6 <> X6) AND ((s6 < 100) OR ((S6 > 99) AND (S6 < 200) AND (mode >= 2)) OR ((S6 > 199) AND (mode = 3))) THEN
    esr_out[cnt] := status_to_ESR(s6, a6, DT_in, TX);
    X6 := S6;
    cnt := cnt + 1;
    esr_flag := TRUE;
  END_IF;
  IF (cnt < 4) AND (s7 <> X7) AND ((s7 < 100) OR ((S7 > 99) AND (S7 < 200) AND (mode >= 2)) OR ((S7 > 199) AND (mode = 3))) THEN
    esr_out[cnt] := status_to_ESR(s7, a7, DT_in, TX);
    X7 := S7;
    cnt := cnt + 1;
    esr_flag := TRUE;
  END_IF;

(* revision history
  hm  26. jan 2007    rev 1.0
    original version

  hm  17. sep 2007  rev 1.1
    replaced time() with T_PLC_MS() for compatibility reasons

  hm  1. dec. 2009  rev 1.2
    changed esr_out to be I/O
*)
END_FUNCTION_BLOCK

(* @PATH := '\/Other' *)
FUNCTION OSCAT_VERSION : DWORD
(*
  oscat_version returns the version number in dword format
  132 is library version 1.32
  if IN = true, the release date will be returned

  version 1.1 16 dec 2007
  programmer  hugo
  tested by   oscat
*)
  VAR_INPUT
    IN : BOOL;
  END_VAR

  IF in THEN
    OSCAT_VERSION := DATE_TO_DWORD(D#2012-01-02);
  ELSE
    OSCAT_VERSION := 333;
  END_IF;

(* revision history
  hm  6. oct 2006 rev 1.0
    original version

  hm  16. dec 2007  rev 1.1
    added possibility to return date and version depending on IN.
*)
END_FUNCTION
